(* IEC 61131-3 sources: daoli-st-library/DL_Process (part 5) *)

(* ---- FB_DL_PackMlUnitMode.st ---- *)
(*
  ==================================================================
  组件名 Component  : FB_DL_PackMlUnitMode
  分类   Category   : DL_Process
  版本   Version    : 1.0.1
  功能   Purpose    : PackML UnitMode 与 PMODE（PackML 状态模型）管理与命令过滤。
                      维护单元模式（生产 / 维护 / 手动 / 换型 / 清洗）与 PackML 状态
                      子集（空闲 / 启动 / 执行 / 保持 / 暂停 / 停止 / 中止 / 清除 /
                      复位 / 完成），按「当前状态 × 当前模式」两张闸对命令做过滤：
                      合法命令被受理并驱动状态迁移，非法命令被拒绝并给出拒绝原因；
                      模式切换仅在空闲 / 停止 / 完成三态允许。
  溯源   Origin     : PackML 状态与 UnitMode 组织为 OMAC PackML 公开标准语义；本件为
                      clean-room 实现，仅借鉴来源分类与参数域组织（来源标签
                      t2-7-packml 的 PackML 状态组织），未复制任何闭源代码行。
  平台   Platform   : 纯 IEC 61131-3（TON / R_TRIG / 枚举比较，无私有库）
  作者   Author     : 道莅代码库 · PLC 编程专家（R55）
  ------------------------------------------------------------------
  边界 Boundary     :
                      一 本件只做模式与状态管理及命令过滤，不执行任何设备动作（属主边界）；
                      二 中止（Abort）与停止（Stop）在全部模式下恒受理（安全侧优先）；
                      三 过渡态（启动 / 保持 / 暂停 / 停止 / 中止 / 清除 / 复位）由外部
                         完成信号 bTransDone 推进，并有过渡超时保护；
                      四 模式切换只在 eIdle / eStopped / eComplete 三态允许，其余态拒绝并留因；
                      五 无全局变量、无外部变量声明、无物理地址寻址。
  输出契约 Output contract:
                      eState / eMode 为锁存状态，只在合法迁移或合法模式切换时改变；
                      bCmdAccepted 为单拍脉冲（内部位置位、统一出口映射后撤销）；
                      eReject 每次拒绝独立留痕，nRejectCnt 饱和累计；
                      eCause 故障级成因与 bError 配对（R45），信息级永不置 bError。
  修订记录 Revision  :
    2026-11-20  v1.0.0  R55 首版（批 4 · 序号 19）
    2026-11-20  v1.0.1  R56 返修（7.5）：段 4 模式受理前补 eModeReq 枚举五选一合法性
                        校验，非法请求改记 eModeBlocked 不采纳（消除一拍非法模式窗口）；
                        段 9 / 段 10 头注释段号回正（原误标 segment 10 / 11）。
  ==================================================================
*)

TYPE E_DL_PmlState :
(
    eIdle        := 0,   // 空闲：允许启动与模式切换 / idle, start and mode change allowed
    eStarting    := 10,  // 启动过渡 / starting transition
    eExecute     := 20,  // 执行 / execute
    eCompleting  := 30,  // 完成过渡 / completing transition
    eComplete    := 40,  // 已完成：允许复位与模式切换 / complete, reset and mode change allowed
    eHolding     := 50,  // 保持过渡 / holding transition
    eHeld        := 60,  // 已保持 / held
    eUnholding   := 70,  // 解除保持过渡 / unholding transition
    eSuspending  := 80,  // 暂停过渡 / suspending transition
    eSuspended   := 90,  // 已暂停 / suspended
    eUnsuspending:= 100, // 解除暂停过渡 / unsuspending transition
    eStopping    := 110, // 停止过渡 / stopping transition
    eStopped     := 120, // 已停止：允许复位与模式切换 / stopped, reset and mode change allowed
    eClearing    := 130, // 清除过渡 / clearing transition
    eAborting    := 140, // 中止过渡 / aborting transition
    eAborted     := 150  // 已中止：只能经清除与复位恢复 / aborted, only clear and reset recover it
);
END_TYPE

TYPE E_DL_UnitMode :
(
    eProduction  := 0,   // 生产模式：全命令集 / production mode with the full command set
    eMaintenance := 10,  // 维护模式：禁暂停 / maintenance mode without suspend
    eManual      := 20,  // 手动模式：禁启动与保持 / manual mode without start and hold
    eChangeover  := 30,  // 换型模式：禁暂停与完成 / changeover mode without suspend and complete
    eCleaning    := 40   // 清洗模式：仅启动 / cleaning mode with start only
);
END_TYPE

TYPE E_DL_PmlCmd :
(
    eNone     := 0,      // 无命令 / no command
    eStart    := 10,     // 启动 / start
    eHold     := 20,     // 保持 / hold
    eUnhold   := 30,     // 解除保持 / unhold
    eSuspend  := 40,     // 暂停 / suspend
    eUnsuspend:= 50,     // 解除暂停 / unsuspend
    eStop     := 60,     // 停止 / stop
    eAbort    := 70,     // 中止 / abort
    eClear    := 80,     // 清除 / clear
    eReset    := 90,     // 复位 / reset
    eComplete := 100     // 完成 / complete
);
END_TYPE

TYPE E_DL_PmlReject :
(
    eNone            := 0, // 无拒绝 / no rejection
    eNoCmd           := 10, // 本拍无命令 / no command in this scan
    eIllegalState    := 20, // 该状态不接受此命令 / the current state does not accept this command
    eModeBlocked     := 30, // 当前模式禁止此命令 / the current mode blocks this command
    eModeLocked      := 40, // 当前状态不允许切换模式 / the current state does not allow a mode change
    eTransTimeout    := 50  // 过渡超时（故障级，与 bError 配对）/ transition timeout, a fault paired with bError
);
END_TYPE

FUNCTION_BLOCK FB_DL_PackMlUnitMode
VAR_INPUT
    bEnable      : BOOL := TRUE;             // 使能，失能时不受理命令并回空闲 [-] / enable, no command is accepted when disabled and the state returns to idle
    bReset       : BOOL := FALSE;           // 复位上升沿清故障锁存并回空闲 [-] / reset rising edge clears the fault latch and returns to idle
    bCmdStrobe   : BOOL := FALSE;            // 命令选通脉冲，上升沿消费 eCmdReq [-] / command strobe, eCmdReq is consumed on the rising edge
    eCmdReq      : E_DL_PmlCmd := E_DL_PmlCmd.eNone;   // 命令请求 [枚举] / requested command [enum]
    bModeStrobe  : BOOL := FALSE;            // 模式切换选通脉冲，上升沿消费 eModeReq [-] / mode change strobe, eModeReq is consumed on the rising edge
    eModeReq     : E_DL_UnitMode := E_DL_UnitMode.eProduction; // 模式请求 [枚举] / requested unit mode [enum]
    bTransDone   : BOOL := FALSE;            // 过渡完成信号（外部动作已完成）[-] / transition done signal from the external action
    tTransTo     : TIME := T#60S;            // 过渡超时 [毫秒]，域 大于零 / transition timeout [millisecond], domain above zero
END_VAR
VAR_OUTPUT
    eState       : E_DL_PmlState := E_DL_PmlState.eIdle;     // PackML 状态出口 [枚举] / PackML state outlet [enum]
    eMode        : E_DL_UnitMode := E_DL_UnitMode.eProduction; // 单元模式出口 [枚举] / unit mode outlet [enum]
    eAccepted    : E_DL_PmlCmd := E_DL_PmlCmd.eNone;         // 最近受理命令 [枚举] / last accepted command [enum]
    eReject      : E_DL_PmlReject := E_DL_PmlReject.eNone;   // 本拍拒绝原因 [枚举] / rejection reason of this scan [enum]
    bCmdAccepted : BOOL := FALSE;            // 命令受理单拍脉冲 [-] / command accepted single-shot pulse
    bModeAllowed : BOOL := FALSE;            // 当前状态是否允许切换模式 [-] / whether the current state allows a mode change
    bTransBusy   : BOOL := FALSE;            // 处于过渡态 [-] / inside a transition state
    uRejectCnt   : UDINT := 0;               // 拒绝计数（饱和到上限）[次] / rejection count, saturated [count]
    eCause       : E_DL_PmlReject := E_DL_PmlReject.eNone;   // 成因出口（复用拒绝枚举，故障级与 bError 配对）/ cause outlet reusing the reject enum, fault grade paired with bError
    bError       : BOOL := FALSE;            // 故障锁存标志 [-] / fault latch flag
END_VAR
VAR
    rtStrobe     : R_TRIG;                   // 命令选通沿检测，段 0 无条件刷新 / command strobe edge detector, refreshed unconditionally in segment zero
    rtMode       : R_TRIG;                   // 模式选通沿检测，段 0 无条件刷新 / mode strobe edge detector, refreshed unconditionally in segment zero
    rtReset      : R_TRIG;                   // 复位沿检测，段 0 无条件刷新 / reset edge detector, refreshed unconditionally in segment zero
    tonTrans     : TON;                      // 过渡超时，段 0 无条件刷新 / transition timeout, refreshed unconditionally in segment zero
    _eState      : E_DL_PmlState := E_DL_PmlState.eIdle;     // 内部状态，CASE 唯一写入目标 / internal state, the only CASE write target
    _eMode       : E_DL_UnitMode := E_DL_UnitMode.eProduction; // 内部模式锁存 / internal mode latch
    _eReject     : E_DL_PmlReject := E_DL_PmlReject.eNone;   // 本拍拒绝原因工作值 / rejection reason working value
    _eAccepted   : E_DL_PmlCmd := E_DL_PmlCmd.eNone;         // 本拍受理命令工作值（出口映射源）[枚举] / accepted command working value, source of the outlet [enum]
    _bFault      : BOOL := FALSE;            // 故障锁存位 [-] / fault latch bit
    _bInit       : BOOL := FALSE;            // 首扫初始化完成标志（R310）/ first scan initialisation flag
    _bAccInt     : BOOL := FALSE;            // 受理脉冲内部位，统一出口映射 / internal accepted bit, mapped at the unified outlet
    _bAccepted   : BOOL := FALSE;            // 本拍是否受理了命令 [-] / whether a command was accepted this scan
    _bTransBusy  : BOOL := FALSE;            // 过渡态判定 [-] / transition state verdict
    _bModeAllowed: BOOL := FALSE;            // 模式切换许可 [-] / mode change permission
    _bAllowStart : BOOL := FALSE;            // 模式允许启动 [-] / the mode allows start
    _bAllowHold  : BOOL := FALSE;            // 模式允许保持 [-] / the mode allows hold
    _bAllowSusp  : BOOL := FALSE;            // 模式允许暂停 [-] / the mode allows suspend
    _bAllowCompl : BOOL := FALSE;            // 模式允许完成 [-] / the mode allows complete
    _bModeValid  : BOOL := FALSE;            // 模式枚举合法 [-] / the mode enumeration is legal
    _bModeReqOk  : BOOL := FALSE;            // 模式请求枚举五选一合法性 [-] / whether the requested mode is one of the five legal members
    _uReject     : UDINT := 0;               // 拒绝计数工作值 [次] / rejection count working value [count]
END_VAR
VAR CONSTANT
    DL_PML_REJ_MAX : UDINT := 2000000000;    // 拒绝计数饱和上限（常量在 DINT 可表范围内）[次] / rejection count saturation ceiling, the constant fits in DINT
END_VAR

// 段 0｜定时器与沿检测无条件周期刷新（禁入分支），IN 只串过渡态闸 / segment 0, unconditional refresh with the transition gate on IN only
rtStrobe(CLK := bCmdStrobe); // 命令选通沿无条件刷新 / unconditional refresh of the command strobe
rtMode(CLK := bModeStrobe); // 模式选通沿无条件刷新 / unconditional refresh of the mode strobe
rtReset(CLK := bReset); // 复位沿无条件刷新 / unconditional refresh of the reset edge
tonTrans(IN := _bTransBusy AND (NOT _bFault) AND bEnable, PT := tTransTo); // 过渡超时，仅在过渡态计时 / transition timeout timing only inside a transition state

// 段 1｜首扫初始化（R310）/ segment 1, first scan initialisation
IF NOT _bInit THEN // 首扫一拍 / the very first scan
    _bInit := TRUE; // 置首扫完成标志 / raise the first scan flag
    _eState := E_DL_PmlState.eIdle; // 状态从空闲起步 / the state starts at idle
    _eMode := E_DL_UnitMode.eProduction; // 模式从生产起步 / the mode starts at production
    _eReject := E_DL_PmlReject.eNone; // 拒绝原因清零 / clear the rejection reason
    _bFault := FALSE; // 故障锁存清零 / clear the fault latch
    _uReject := 0; // 拒绝计数清零 / clear the rejection count
END_IF

// 段 2｜复位沿作用域：清锁存 / 迁状态 / 清脉冲内部位（模式保持，避免复位改工艺模式）/ segment 2, reset edge scope
IF rtReset.Q THEN // 复位沿 / reset edge
    _bFault := FALSE; // 作用域一：清故障锁存 / scope one, clear the fault latch
    _eReject := E_DL_PmlReject.eNone; // 作用域一：清拒绝原因 / scope one, clear the rejection reason
    _eState := E_DL_PmlState.eIdle; // 作用域二：迁回空闲 / scope two, migrate back to idle
    _bAccInt := FALSE; // 作用域二：清受理脉冲内部位 / scope two, clear the internal accepted bit
END_IF

// 段 3｜模式合法性与模式命令白名单（模式闸） / segment 3, mode validity and the per mode command whitelist
_bModeValid := (_eMode = E_DL_UnitMode.eProduction) OR (_eMode = E_DL_UnitMode.eMaintenance) OR (_eMode = E_DL_UnitMode.eManual) OR (_eMode = E_DL_UnitMode.eChangeover) OR (_eMode = E_DL_UnitMode.eCleaning); // 模式枚举五选一 / the mode is one of five
IF NOT _bModeValid THEN // 模式非法 / the mode is illegal
    _eMode := E_DL_UnitMode.eProduction; // 两级回退（R117）：一级回生产模式 / stage one of the two stage fallback, back to production
END_IF
_bAllowStart := (_eMode = E_DL_UnitMode.eProduction) OR (_eMode = E_DL_UnitMode.eMaintenance) OR (_eMode = E_DL_UnitMode.eChangeover) OR (_eMode = E_DL_UnitMode.eCleaning); // 启动白名单：手动模式禁启动 / start whitelist, manual mode forbids start
_bAllowHold := (_eMode = E_DL_UnitMode.eProduction) OR (_eMode = E_DL_UnitMode.eMaintenance) OR (_eMode = E_DL_UnitMode.eChangeover); // 保持白名单：手动与清洗禁保持 / hold whitelist, manual and cleaning forbid hold
_bAllowSusp := (_eMode = E_DL_UnitMode.eProduction); // 暂停白名单：仅生产模式 / suspend whitelist, production only
_bAllowCompl := (_eMode = E_DL_UnitMode.eProduction); // 完成白名单：仅生产模式 / complete whitelist, production only
_bModeAllowed := (_eState = E_DL_PmlState.eIdle) OR (_eState = E_DL_PmlState.eStopped) OR (_eState = E_DL_PmlState.eComplete); // 模式切换许可：空闲 / 停止 / 完成三态 / mode change allowed in idle, stopped and complete only

// 段 4｜模式切换：许可态内受理，非许可态留拒绝原因 / segment 4, mode change acceptance with a rejection trail
_eReject := E_DL_PmlReject.eNone; // 本拍拒绝原因预置空 / preset the rejection reason to none
_bModeReqOk := (eModeReq = E_DL_UnitMode.eProduction) OR (eModeReq = E_DL_UnitMode.eMaintenance) OR (eModeReq = E_DL_UnitMode.eManual) OR (eModeReq = E_DL_UnitMode.eChangeover) OR (eModeReq = E_DL_UnitMode.eCleaning); // 模式请求枚举五选一判式（R56 返修补齐）/ the requested mode is one of five legal members
IF rtMode.Q THEN // 模式选通沿 / mode strobe edge
    IF NOT bEnable THEN // 失能 / disabled
        _eReject := E_DL_PmlReject.eModeLocked; // 拒绝原因：失能不受理 / rejection reason, disabled
    ELSIF NOT _bModeReqOk THEN // 模式请求枚举非法 / the requested mode is illegal
        _eReject := E_DL_PmlReject.eModeBlocked; // 拒绝原因：非法模式请求不采纳（R56 返修补齐，消除一拍非法模式窗口）/ rejection reason, an illegal mode request is not adopted
    ELSIF _bModeAllowed THEN // 许可态 / inside a permitted state
        _eMode := eModeReq; // 采纳请求模式 / adopt the requested mode
    ELSE // 非许可态 / outside a permitted state
        _eReject := E_DL_PmlReject.eModeLocked; // 拒绝原因：状态锁模式 / rejection reason, the state locks the mode
    END_IF
END_IF

// 段 5｜过渡态判定 / segment 5, transition state verdict
_bTransBusy := (_eState = E_DL_PmlState.eStarting) OR (_eState = E_DL_PmlState.eCompleting) OR (_eState = E_DL_PmlState.eHolding) OR (_eState = E_DL_PmlState.eUnholding) OR (_eState = E_DL_PmlState.eSuspending) OR (_eState = E_DL_PmlState.eUnsuspending) OR (_eState = E_DL_PmlState.eStopping) OR (_eState = E_DL_PmlState.eClearing) OR (_eState = E_DL_PmlState.eAborting); // 九个过渡态之一 / one of the nine transition states

// 段 6｜过渡推进：外部完成信号或过渡超时（超时即中止并留故障级原因）/ segment 6, transition advancement by the external signal or by a timeout
IF _bTransBusy THEN // 过渡态内 / inside a transition state
    IF bTransDone THEN // 外部动作完成 / the external action completed
        CASE _eState OF
        E_DL_PmlState.eStarting: // 启动过渡完成 / starting completed
            _eState := E_DL_PmlState.eExecute; // 进执行态 / enter execute
        E_DL_PmlState.eCompleting: // 完成过渡完成 / completing completed
            _eState := E_DL_PmlState.eComplete; // 进已完成态 / enter complete
        E_DL_PmlState.eHolding: // 保持过渡完成 / holding completed
            _eState := E_DL_PmlState.eHeld; // 进已保持态 / enter held
        E_DL_PmlState.eUnholding: // 解除保持过渡完成 / unholding completed
            _eState := E_DL_PmlState.eExecute; // 回执行态 / back to execute
        E_DL_PmlState.eSuspending: // 暂停过渡完成 / suspending completed
            _eState := E_DL_PmlState.eSuspended; // 进已暂停态 / enter suspended
        E_DL_PmlState.eUnsuspending: // 解除暂停过渡完成 / unsuspending completed
            _eState := E_DL_PmlState.eExecute; // 回执行态 / back to execute
        E_DL_PmlState.eStopping: // 停止过渡完成 / stopping completed
            _eState := E_DL_PmlState.eStopped; // 进已停止态 / enter stopped
        E_DL_PmlState.eClearing: // 清除过渡完成 / clearing completed
            _eState := E_DL_PmlState.eIdle; // 回空闲态 / back to idle
        E_DL_PmlState.eAborting: // 中止过渡完成 / aborting completed
            _eState := E_DL_PmlState.eAborted; // 进已中止态 / enter aborted
        ELSE // 非法过渡态兜底（R128）/ illegal transition fallback
            _eState := E_DL_PmlState.eIdle; // 回空闲态 / back to idle
        END_CASE
    ELSIF tonTrans.Q THEN // 过渡超时 / the transition timed out
        _eReject := E_DL_PmlReject.eTransTimeout; // 故障级原因（与 bError 配对，R45）/ fault grade reason paired with bError
        _bFault := TRUE; // 置故障锁存 / raise the fault latch
        _eState := E_DL_PmlState.eAborting; // 强制走中止过渡 / force the aborting transition
    END_IF
END_IF

// 段 7｜命令过滤：状态闸在前、模式闸在后，两闸顺序固定（先判状态可接受性，再判模式白名单）/ segment 7, command filtering with the state gate before the mode gate
_eAccepted := E_DL_PmlCmd.eNone; // 受理命令预置空 / preset the accepted command to none
_bAccepted := FALSE; // 受理标志预置假 / preset the accepted flag to false
IF rtStrobe.Q AND bEnable AND (NOT _bFault) AND (NOT _bTransBusy) THEN // 选通沿、使能、无故障、非过渡态 / strobe while enabled, unfaulted and outside a transition
    IF eCmdReq = E_DL_PmlCmd.eNone THEN // 无命令 / no command
        _eReject := E_DL_PmlReject.eNoCmd; // 拒绝原因：无命令 / rejection reason, no command
    ELSE
        // 段 7.1｜状态闸：按当前状态给出可接受的命令集合 / segment 7.1, the state gate defines the acceptable command set
        CASE _eState OF
        E_DL_PmlState.eIdle: // 空闲态：启动 / 中止 / 复位 / 清除 / 模式许可 / idle state
            IF eCmdReq = E_DL_PmlCmd.eStart THEN // 启动 / start
                IF _bAllowStart THEN // 模式允许 / the mode allows it
                    _eState := E_DL_PmlState.eStarting; // 迁启动过渡 / enter starting
                    _eAccepted := E_DL_PmlCmd.eStart; // 受理启动 / accept start
                    _bAccepted := TRUE; // 置受理标志 / raise the accepted flag
                ELSE
                    _eReject := E_DL_PmlReject.eModeBlocked; // 模式闸拒绝 / blocked by the mode gate
                END_IF
            ELSIF eCmdReq = E_DL_PmlCmd.eAbort THEN // 中止 / abort
                _eState := E_DL_PmlState.eAborting; // 迁中止过渡 / enter aborting
                _eAccepted := E_DL_PmlCmd.eAbort; // 受理中止 / accept abort
                _bAccepted := TRUE; // 置受理标志 / raise the accepted flag
            ELSIF eCmdReq = E_DL_PmlCmd.eReset THEN // 复位 / reset
                _eState := E_DL_PmlState.eClearing; // 空闲态的复位等价于清除 / a reset from idle behaves as clearing
                _eAccepted := E_DL_PmlCmd.eReset; // 受理复位 / accept reset
                _bAccepted := TRUE; // 置受理标志 / raise the accepted flag
            ELSIF eCmdReq = E_DL_PmlCmd.eClear THEN // 清除 / clear
                _eState := E_DL_PmlState.eClearing; // 迁清除过渡 / enter clearing
                _eAccepted := E_DL_PmlCmd.eClear; // 受理清除 / accept clearing
                _bAccepted := TRUE; // 置受理标志 / raise the accepted flag
            ELSE // 其它命令 / any other command
                _eReject := E_DL_PmlReject.eIllegalState; // 状态闸拒绝 / blocked by the state gate
            END_IF
        E_DL_PmlState.eExecute: // 执行态：保持 / 暂停 / 停止 / 完成 / 中止 / execute state
            IF eCmdReq = E_DL_PmlCmd.eHold THEN // 保持 / hold
                IF _bAllowHold THEN // 模式允许 / the mode allows it
                    _eState := E_DL_PmlState.eHolding; // 迁保持过渡 / enter holding
                    _eAccepted := E_DL_PmlCmd.eHold; // 受理保持 / accept hold
                    _bAccepted := TRUE; // 置受理标志 / raise the accepted flag
                ELSE
                    _eReject := E_DL_PmlReject.eModeBlocked; // 模式闸拒绝 / blocked by the mode gate
                END_IF
            ELSIF eCmdReq = E_DL_PmlCmd.eSuspend THEN // 暂停 / suspend
                IF _bAllowSusp THEN // 模式允许 / the mode allows it
                    _eState := E_DL_PmlState.eSuspending; // 迁暂停过渡 / enter suspending
                    _eAccepted := E_DL_PmlCmd.eSuspend; // 受理暂停 / accept suspend
                    _bAccepted := TRUE; // 置受理标志 / raise the accepted flag
                ELSE
                    _eReject := E_DL_PmlReject.eModeBlocked; // 模式闸拒绝 / blocked by the mode gate
                END_IF
            ELSIF eCmdReq = E_DL_PmlCmd.eComplete THEN // 完成 / complete
                IF _bAllowCompl THEN // 模式允许 / the mode allows it
                    _eState := E_DL_PmlState.eCompleting; // 迁完成过渡 / enter completing
                    _eAccepted := E_DL_PmlCmd.eComplete; // 受理完成 / accept complete
                    _bAccepted := TRUE; // 置受理标志 / raise the accepted flag
                ELSE
                    _eReject := E_DL_PmlReject.eModeBlocked; // 模式闸拒绝 / blocked by the mode gate
                END_IF
            ELSIF eCmdReq = E_DL_PmlCmd.eStop THEN // 停止（安全侧恒受理）/ stop, always accepted on the safety side
                _eState := E_DL_PmlState.eStopping; // 迁停止过渡 / enter stopping
                _eAccepted := E_DL_PmlCmd.eStop; // 受理停止 / accept stop
                _bAccepted := TRUE; // 置受理标志 / raise the accepted flag
            ELSIF eCmdReq = E_DL_PmlCmd.eAbort THEN // 中止（安全侧恒受理）/ abort, always accepted
                _eState := E_DL_PmlState.eAborting; // 迁中止过渡 / enter aborting
                _eAccepted := E_DL_PmlCmd.eAbort; // 受理中止 / accept abort
                _bAccepted := TRUE; // 置受理标志 / raise the accepted flag
            ELSE // 其它命令 / any other command
                _eReject := E_DL_PmlReject.eIllegalState; // 状态闸拒绝 / blocked by the state gate
            END_IF
        E_DL_PmlState.eHeld: // 已保持态：解除保持 / 停止 / 中止 / held state
            IF eCmdReq = E_DL_PmlCmd.eUnhold THEN // 解除保持 / unhold
                _eState := E_DL_PmlState.eUnholding; // 迁解除保持过渡 / enter unholding
                _eAccepted := E_DL_PmlCmd.eUnhold; // 受理解除保持 / accept unhold
                _bAccepted := TRUE; // 置受理标志 / raise the accepted flag
            ELSIF eCmdReq = E_DL_PmlCmd.eStop THEN // 停止 / stop
                _eState := E_DL_PmlState.eStopping; // 迁停止过渡 / enter stopping
                _eAccepted := E_DL_PmlCmd.eStop; // 受理停止 / accept stop
                _bAccepted := TRUE; // 置受理标志 / raise the accepted flag
            ELSIF eCmdReq = E_DL_PmlCmd.eAbort THEN // 中止 / abort
                _eState := E_DL_PmlState.eAborting; // 迁中止过渡 / enter aborting
                _eAccepted := E_DL_PmlCmd.eAbort; // 受理中止 / accept abort
                _bAccepted := TRUE; // 置受理标志 / raise the accepted flag
            ELSE // 其它命令 / any other command
                _eReject := E_DL_PmlReject.eIllegalState; // 状态闸拒绝 / blocked by the state gate
            END_IF
        E_DL_PmlState.eSuspended: // 已暂停态：解除暂停 / 停止 / 中止 / suspended state
            IF eCmdReq = E_DL_PmlCmd.eUnsuspend THEN // 解除暂停 / unsuspend
                _eState := E_DL_PmlState.eUnsuspending; // 迁解除暂停过渡 / enter unsuspending
                _eAccepted := E_DL_PmlCmd.eUnsuspend; // 受理解除暂停 / accept unsuspend
                _bAccepted := TRUE; // 置受理标志 / raise the accepted flag
            ELSIF eCmdReq = E_DL_PmlCmd.eStop THEN // 停止 / stop
                _eState := E_DL_PmlState.eStopping; // 迁停止过渡 / enter stopping
                _eAccepted := E_DL_PmlCmd.eStop; // 受理停止 / accept stop
                _bAccepted := TRUE; // 置受理标志 / raise the accepted flag
            ELSIF eCmdReq = E_DL_PmlCmd.eAbort THEN // 中止 / abort
                _eState := E_DL_PmlState.eAborting; // 迁中止过渡 / enter aborting
                _eAccepted := E_DL_PmlCmd.eAbort; // 受理中止 / accept abort
                _bAccepted := TRUE; // 置受理标志 / raise the accepted flag
            ELSE // 其它命令 / any other command
                _eReject := E_DL_PmlReject.eIllegalState; // 状态闸拒绝 / blocked by the state gate
            END_IF
        E_DL_PmlState.eComplete: // 已完成态：复位 / 停止 / 中止 / complete state
            IF (eCmdReq = E_DL_PmlCmd.eReset) OR (eCmdReq = E_DL_PmlCmd.eClear) THEN // 复位或清除 / reset or clear
                _eState := E_DL_PmlState.eClearing; // 迁清除过渡 / enter clearing
                _eAccepted := eCmdReq; // 受理该命令 / accept that command
                _bAccepted := TRUE; // 置受理标志 / raise the accepted flag
            ELSIF eCmdReq = E_DL_PmlCmd.eAbort THEN // 中止 / abort
                _eState := E_DL_PmlState.eAborting; // 迁中止过渡 / enter aborting
                _eAccepted := E_DL_PmlCmd.eAbort; // 受理中止 / accept abort
                _bAccepted := TRUE; // 置受理标志 / raise the accepted flag
            ELSE // 其它命令 / any other command
                _eReject := E_DL_PmlReject.eIllegalState; // 状态闸拒绝 / blocked by the state gate
            END_IF
        E_DL_PmlState.eStopped: // 已停止态：复位 / 清除 / 中止 / stopped state
            IF (eCmdReq = E_DL_PmlCmd.eReset) OR (eCmdReq = E_DL_PmlCmd.eClear) THEN // 复位或清除 / reset or clear
                _eState := E_DL_PmlState.eClearing; // 迁清除过渡 / enter clearing
                _eAccepted := eCmdReq; // 受理该命令 / accept that command
                _bAccepted := TRUE; // 置受理标志 / raise the accepted flag
            ELSIF eCmdReq = E_DL_PmlCmd.eAbort THEN // 中止 / abort
                _eState := E_DL_PmlState.eAborting; // 迁中止过渡 / enter aborting
                _eAccepted := E_DL_PmlCmd.eAbort; // 受理中止 / accept abort
                _bAccepted := TRUE; // 置受理标志 / raise the accepted flag
            ELSE // 其它命令 / any other command
                _eReject := E_DL_PmlReject.eIllegalState; // 状态闸拒绝 / blocked by the state gate
            END_IF
        E_DL_PmlState.eAborted: // 已中止态：只能清除后复位 / aborted state, clear then reset only
            IF eCmdReq = E_DL_PmlCmd.eClear THEN // 清除 / clear
                _eState := E_DL_PmlState.eClearing; // 迁清除过渡 / enter clearing
                _eAccepted := E_DL_PmlCmd.eClear; // 受理清除 / accept clearing
                _bAccepted := TRUE; // 置受理标志 / raise the accepted flag
            ELSE // 其它命令 / any other command
                _eReject := E_DL_PmlReject.eIllegalState; // 状态闸拒绝 / blocked by the state gate
            END_IF
        ELSE // 过渡态不接受新命令 / transition states reject new commands
            _eReject := E_DL_PmlReject.eIllegalState; // 状态闸拒绝 / blocked by the state gate
        END_CASE
    END_IF
ELSIF rtStrobe.Q THEN // 有选通但使能 / 故障 / 过渡态不满足 / a strobe arrived under a blocking condition
    _eReject := E_DL_PmlReject.eIllegalState; // 拒绝原因：条件不满足 / rejection reason, the condition is not met
END_IF

// 段 8｜拒绝计数与受理脉冲内部位 / segment 8, rejection counting and the internal accepted bit
IF NOT (_eReject = E_DL_PmlReject.eNone) THEN // 本拍存在拒绝 / a rejection occurred
    IF _uReject < DL_PML_REJ_MAX THEN // 未达饱和上限 / below the ceiling
        _uReject := _uReject + 1; // 拒绝计数递增 / increment the rejection count
    END_IF
END_IF
IF _bAccepted THEN // 本拍受理了命令 / a command was accepted
    _bAccInt := TRUE; // 受理脉冲内部位置位（统一出口映射，R187）/ raise the internal accepted bit, mapped at the unified outlet
END_IF

// 段 9｜失能语义：不受理命令，状态保持但过渡计时停摆（R191 显式声明）/ segment 9, disabled semantics
IF NOT bEnable THEN // 失能 / disabled
    _bAccInt := FALSE; // 撤受理脉冲内部位 / withdraw the internal accepted bit
    _eReject := E_DL_PmlReject.eModeLocked; // 拒绝原因记模式锁（失能态不支持任何命令）/ rejection reason, disabled blocks every command
END_IF

// 段 10｜统一出口 / segment 10, unified outlet
eState := _eState; // 状态出口单点映射 / single-point state outlet mapping
eMode := _eMode; // 模式出口（锁存量）/ mode outlet from the latch
eAccepted := _eAccepted; // 受理命令出口 / accepted command outlet
eReject := _eReject; // 拒绝原因出口 / rejection reason outlet
bCmdAccepted := _bAccInt; // 受理脉冲映射本拍值 / map the accepted pulse for this scan
_bAccInt := FALSE; // 映射后立即撤销，保证单拍宽度（R187 两段式）/ revoke right after mapping to keep a single-scan width
bModeAllowed := _bModeAllowed; // 模式切换许可出口 / mode change permission outlet
bTransBusy := _bTransBusy; // 过渡态出口 / transition state outlet
uRejectCnt := _uReject; // 拒绝计数出口 / rejection count outlet
eCause := _eReject; // 成因出口与拒绝原因同源（名实双出口，R191）/ the cause outlet shares the rejection source
bError := _bFault; // 故障标志与锁存位同源 / the fault flag shares the latch source
END_FUNCTION_BLOCK

(* ---- FB_DL_PollTempBank.st ---- *)
(*==============================================================================
 * 组件名称 (Component)  : FB_DL_PollTempBank
 * 所属子库 (Sublibrary) : DL_Process
 * 当前版本 (Version)    : 1.0.0
 * 组件分类 (Category)   : 功能块（FUNCTION_BLOCK）· 工艺采集 · 温控器轮询采集行
 * 兼容性   (Platform)   : CODESYS 3.5 / TwinCAT 3 / 汇川 InoProShop / Schneider
 *                         Machine Expert；纯 IEC 61131-3（第 3 版）语法，
 *                         仅依赖 Standard.library（R_TRIG）
 * 功能描述 (Function)   : 一条温控器采集行——对最多 8 台温控器轮询采集过程值与设定值，
 *                         做工程量换算、有效域判定、滑动均值、偏差与最差通道定位，
 *                         输出通道质量掩码与在线台数，连续失败通道自动摘除并自动恢复。
 * 分层声明 (Layering)   : ① 调度归既有轮询主站件（本件内嵌其一个实例，只注入站表与
 *                         节拍参数，不重写调度、重试与超时逻辑）；② 滤波归既有滑动均值件
 *                         （本件为八个通道各持一个实例，只给样本与采样允许）；
 *                         ③ 本件只做「行级编排加通道质量」，不做温控闭环——设定值下发、
 *                         自整定、超温切断属温控器内部或工艺层职责，本件只读不写。
 * 传输层说明 (Transport) : 内嵌的调度实例以库内基类形态声明，其帧收发为抽象桩。生产部署
 *                         时必须由具备真实串口或网口收发的派生块替换该声明，否则调度层会
 *                         锁「传输层未实现」故障、全部通道因轮询不成功而逐台摘除。这一
 *                         失败是**可观测的显式失败**（质量掩码全置位、在线台数为零），
 *                         不会静默给出假温度，故不在本件内把它翻译成故障码。
 * 保持策略 (Hold)       : 坏通道的温度保持上次有效值并在质量掩码里标记，**绝不**用零或
 *                         上限值填充——零摄氏度在锂电烘箱、冷库等场景是合法工况值，用零
 *                         填充会掩盖真实故障（与既有温度扫描件同一纪律）。
 * 摘除与恢复 (Drop)     : 连续失败达到阈值即摘除并置信息码；摘除后仍继续轮询该通道，
 *                         连续两拍有效即自动恢复。若不继续轮询，被摘除的通道永远拿不到
 *                         有效数据、也就永远无法恢复，这是摘除策略必须配对的另一半。
 * 职责边界 (Scope)      : 不做写设定值（只采集）、不做地址表编辑器的校验（站表按默认值
 *                         填充，机型差异由调用方改表）、不做历史归档与报警分级。
 * 开源溯源 (Origin)     : 来源标签 roadmap-p0 加 t1-4。原创实现（参考 ROADMAP §13.6 P0
 *                         条目「温控器轮询采集行（复用轮询主站与滑动均值）」的需求定义，
 *                         以及 CODESYS Forge ModbusFB 族「调度与传输分层」的组织方式）。
 *                         仅借组织方式与参数域，编排逻辑、通道质量掩码、摘除与恢复策略、
 *                         枚举、状态机与全部码位 100% 本库独立设计，clean-room 实现，
 *                         不复制任何示例代码与注释。
 * 依赖     (Depends)    : ST_DL_PollItem 与 FB_DL_ModbusPollMaster（DL_Process 既有件，
 *                         本件只引用不声明）；FB_DL_MovingAverage（DL_MathData 既有件）；
 *                         Standard.library: R_TRIG
 * 故障码表 (Error codes):
 *   16#0005_0108【信息级】台数、窗口长度或摘除阈值越界已钳位
 *   16#0005_0109【信息级】通道连续失败达到阈值已摘除（仍继续轮询以便自动恢复）
 *   16#0005_010A【信息级】滤波窗口为 1，均值等于瞬时值（无滤波能力）
 *   16#0005_0207【故障级】换算比例非正，量纲错且含零乘隐患（锁存）
 *   16#0005_0208【故障级】有效温度域为空，任何读数都会被判无效（锁存）
 *   16#0005_0209【故障级】非法状态兜底（锁存，终端安全态）
 * 码位占用 (Slot)       : 信息级 0108 / 0109 / 010A；故障级 0207 / 0208 / 0209。
 *                         全部落在 R12 本件分配块内，无跨块借用、无段外哨兵值。
 * 拍序纪律 (Cycle order) :
 *   ① ePhase        ：段 7 状态机（唯一位移点），段 8 复位分支是唯一回退点
 *   ② 三个生效参数   ：段 4 单点钳位，后续所有数组访问与循环上限都取这三个生效值
 *   ③ 质量掩码       ：段 6 装配后整值写出，与本拍在线台数、最差通道同拍一致
 *   ④ uErrorId       ：段 9 单一优先级链，全拍只写一次
 * 验收向量 (Acceptance) :
 *   V1 单台正常：台数 1、过程值 253、设定值 250、比例 0.1 → 温度 25.3、设定 25.0、
 *      偏差 0.3、质量掩码为零、在线 1 台
 *   V2 超域：第 2 台过程值 3200（换算 320.0 高于上限 200）→ 该通道无效、温度保持、
 *      质量掩码位 1 置位、连续失败计数 1
 *   V3 摘除：第 3 台连续三拍轮询失败、阈值为 3 → 第 3 拍摘除、质量掩码位 2 置位、
 *      在线台数减 1、码 0109
 *   V4 最差通道：两通道偏差分别负 3.5 与正 4.2 → 最差通道号为 4、最差偏差正 4.2
 *   V5 量纲错：比例为 0 → 故障位置位、码 0207、各通道温度保持
 * 偏离留档 (Deviation)  :
 *   ① 规格第 3.18 节正文提到「评估相」，但 §2.1 的枚举只有三成员。本件按枚举实现，
 *      把逐通道评估并入轮询相的固定段完成，不新增枚举成员，避免枚举与码表、文档三处
 *      不一致。
 *   ② 规格要求「内嵌调度实例」，但库内调度基类的传输层为抽象桩，无法在本文件内以派生块
 *      替换其声明。本件保留基类实例并在头注释写明部署要求，把「传输层未就绪」表现为
 *      质量掩码全坏这一可观测结果，而不是伪造成功。
 *   ③ 参数钳位放在状态机之前的固定段（而非待机相），理由：台数决定站表填充与循环上限，
 *      必须每拍先于任何数组访问生效，否则上电首拍会用未钳位值访问数组。
 * 修订历史 (Revision)   :
 *   2026-11-15  v1.0.0  首版落盘（R12 · 泳道 C · 温控器轮询采集行 P0 件）
 *============================================================================*)

(*------------------------------------------------------------------------------
 * 枚举: E_DL_TempBankPhase（本块相位，归属本功能块并同文件发布）
 *       Phase enumeration owned by this block
 *-----------------------------------------------------------------------------*)
TYPE E_DL_TempBankPhase :
(
    eIdle    := 0,   // 待机：未使能或参数闸门未过，输出保持 / Idle, disabled or the gate has not passed
    ePolling := 10,  // 轮询：调度实例推进轮询，同时做逐通道换算与质量判定 / Polling with per-channel evaluation
    eFault   := 99   // 故障：量纲错、有效域为空或非法状态，需复位退出 / Fault, needs a reset to leave
);
END_TYPE

FUNCTION_BLOCK FB_DL_PollTempBank
VAR_INPUT
    bEnable        : BOOL;                              // 使能，FALSE 时暂停轮询并保持输出 [-] / Enable, polling paused and outputs held while FALSE
    bReset         : BOOL;                              // 复位故障与摘除状态，上升沿有效 [-] / Rising edge clears the fault and the drop state
    nDeviceCount   : INT := 4;                          // 温控器台数 [台]，有效域 1 到 8 / Device count, one to eight
    anSlaveAddr    : ARRAY[1..8] OF USINT;              // 各台从站地址 [1 到 247] / Slave address per device
    auPvRaw        : ARRAY[1..8] OF INT;                // 各台过程值原始寄存器，由传输层写入 [原始码] / Raw process values written by the transport
    auSvRaw        : ARRAY[1..8] OF INT;                // 各台设定值原始寄存器 [原始码] / Raw setpoints
    abPollOk       : ARRAY[1..8] OF BOOL;               // 各台本次轮询成功标志 [-] / Per-device poll success flags
    fScaleGain     : REAL := 0.1;                       // 原始码到温度的比例 [摄氏度每码]，域大于 0 / Raw to temperature gain, must exceed zero
    fScaleOffset   : REAL := 0.0;                       // 零点偏移 [摄氏度] / Zero offset in degrees Celsius
    fRangeMin      : REAL := -50.0;                     // 有效温度下限 [摄氏度] / Valid temperature lower bound
    fRangeMax      : REAL := 200.0;                     // 有效温度上限 [摄氏度] / Valid temperature upper bound
    nFilterLen     : INT := 8;                          // 滑动均值窗口长度 [拍]，有效域 1 到 32 / Moving average window, one to thirty-two
    nDropAfterFails: INT := 3;                          // 连续失败多少次摘除通道 [次]，有效域 1 到 10 / Failures before dropping a channel
END_VAR
VAR_OUTPUT
    afTempC        : ARRAY[1..8] OF REAL;               // 各台温度 [摄氏度]，坏通道保持上次有效值 / Temperature per device, bad channels hold the last value
    afSetpointC    : ARRAY[1..8] OF REAL;               // 各台设定值 [摄氏度] / Setpoint per device
    afDeviation    : ARRAY[1..8] OF REAL;               // 各台偏差，过程值减设定值 [摄氏度] / Deviation, process minus setpoint
    afTempAvg      : ARRAY[1..8] OF REAL;               // 各台滑动均值 [摄氏度] / Per-device moving average
    auCommFailCnt  : ARRAY[1..8] OF UINT;               // 各台连续失败次数，饱和到上限 [次] / Consecutive failure counter per device, saturated
    uQualityMask   : WORD;                              // 通道坏质量掩码，位 n 减一 对应第 n 台 [位串] / Bad channel mask, bit n minus one is device n
    nOnlineCount   : INT;                               // 在线台数 [台] / Online device count
    nWorstIdx      : INT;                               // 偏差绝对值最大的在线通道号，0 表示无 [通道号] / Channel with the largest absolute deviation
    fWorstDev      : REAL;                              // 该通道的有符号偏差值 [摄氏度] / Signed deviation of that channel
    bError         : BOOL;                              // 故障级锁存，仅 0207 至 0209 置位 [-] / Latched fault, only fault level codes set it
    uErrorId       : UDINT;                             // 事件码，0 表示无事件 [代码] / Event code, zero means none
    eState         : E_DL_TempBankPhase;                // 主状态机当前相位 [-] / Current phase of the main state machine
END_VAR
VAR_IN_OUT
    aPollTable     : ARRAY[0..15] OF ST_DL_PollItem;    // 轮询站表，由内嵌调度实例持有并更新统计 [-] / Poll table owned by the embedded scheduler
END_VAR
VAR
    fbPoll         : FB_DL_ModbusPollMaster;            // 内嵌轮询调度实例，主周期无条件调用 / Embedded poll scheduler, called unconditionally
    afbAvg         : ARRAY[1..8] OF FB_DL_MovingAverage; // 逐通道滑动均值实例，主周期无条件全量调用 / Per-channel moving average instances
    fbTrigReset    : R_TRIG;                            // 复位沿检测，主周期无条件刷新 [-] / Reset edge detector, refreshed unconditionally
    ePhase         : E_DL_TempBankPhase := E_DL_TempBankPhase.eIdle; // 内部相位，对外经 eState 输出 [-] / Internal phase exported as eState
    bInit          : BOOL := FALSE;                     // 首扫标志，初值 FALSE，判据取非 [-] / First-scan flag initialised FALSE
    bFaultLatch    : BOOL;                              // 故障锁存，仅复位分支清除 [-] / Fault latch, cleared by the reset path only
    uErrInt        : UDINT;                             // 故障级码寄存，锁存型 [代码] / Latched fault level code register
    uInfoCode      : UDINT;                             // 本拍信息级码，每拍重算 [代码] / Info level code recomputed every scan
    nDevUse        : INT := 1;                          // 生效台数，钳位后 [台] / Effective device count after clamping
    nFilterUse     : INT := 1;                          // 生效窗口长度，钳位后 [拍] / Effective window length after clamping
    nDropUse       : INT := 1;                          // 生效摘除阈值，钳位后 [次] / Effective drop threshold after clamping
    fGainUse       : REAL := 1.0;                       // 生效换算比例 [摄氏度每码] / Effective gain
    bEval          : BOOL;                              // 本拍执行通道评估 [-] / Evaluation enabled flag of this scan
    bDropEvent     : BOOL;                              // 本拍有通道被摘除 [-] / A channel was dropped this scan
    fVal           : REAL;                              // 单通道温度 [摄氏度] / Single channel temperature
    fSp            : REAL;                              // 单通道设定值 [摄氏度] / Single channel setpoint
    fDevAbs        : REAL;                              // 偏差绝对值 [摄氏度] / Absolute deviation
    fWorstTmp      : REAL;                              // 最差偏差绝对值暂存 [摄氏度] / Worst absolute deviation temporary
    uQBuild        : WORD;                              // 质量掩码装配 [位串] / Quality mask under assembly
    nOnline        : INT;                               // 在线计数 [台] / Online counter
    nWorst         : INT;                               // 最差通道号 [通道号] / Worst channel number
    abOkTmp        : ARRAY[1..8] OF BOOL;               // 各通道本拍有效标志 [-] / Per-channel validity of this scan
    abDropped      : ARRAY[1..8] OF BOOL;               // 通道已摘除标志 [-] / Channel dropped flags
    anRecover      : ARRAY[1..8] OF INT;                // 摘除后连续有效拍数 [拍] / Consecutive valid scans after a drop
    bValFin        : BOOL;                              // 换算值有限标志 [-] / Finite converted value flag
    nGuard         : DINT;                              // 循环守卫计数 [次]，上限常量化 / Loop guard counter with a constant bound
    i              : INT;                               // 通道索引 [1..8] / Channel loop index
    k              : INT;                               // 站表索引 [0..15] / Poll table loop index
END_VAR
VAR CONSTANT
    DL_DEV_MAX     : INT := 8;                          // 温控器台数上限 [台] / Device count limit
    DL_FILT_MAX    : INT := 32;                         // 滤波窗口上限 [拍] / Window length limit
    DL_DROP_MAX    : INT := 10;                         // 摘除阈值上限 [次] / Drop threshold limit
    DL_TABLE_MAX   : INT := 16;                         // 站表长度 [项] / Poll table length
    DL_FAIL_MAX    : UINT := 9999;                      // 连续失败计数饱和值 [次] / Failure counter saturation
    DL_MASK_ONE    : WORD := 16#0001;                   // 单通道基准位 [位串] / Single channel base bit
    DL_MASK_NONE   : WORD := 16#0000;                   // 全零掩码基准 [位串] / All zero mask reference
    DL_GAIN_MIN    : REAL := 1.0E-6;                    // 比例最小正值 [摄氏度每码] / Minimum positive gain
    DL_GAIN_SAFE   : REAL := 1.0;                       // 比例非法时的兜底值 [摄氏度每码] / Safe gain used when the input is illegal
    DL_TEMP_MAX    : REAL := 1.0E6;                     // 温度量级上限，超出视为非有限 [摄氏度] / Temperature magnitude bound
    DL_GUARD_MAX   : DINT := 64;                        // 循环守卫上限 [次] / Loop guard bound
    DL_RECOVER_NEED: INT := 2;                          // 自动恢复所需的连续有效拍数 [拍] / Valid scans required for an automatic recovery
    DL_FUNC_READ   : USINT := 3;                        // 读保持寄存器功能码 [功能码] / Read holding registers function code
    DL_REG_QTY     : UINT := 2;                         // 每站连续读两个寄存器，过程值与设定值 [个] / Two registers per station
    DL_REG_START   : UINT := 0;                         // 站表起始地址 [寄存器地址] / Station start address
    DL_RESP_TO     : TIME := T#500MS;                   // 单事务响应超时 [毫秒] / Per-transaction response timeout
    DL_POLL_GAP    : TIME := T#50MS;                    // 相邻事务最小间隔 [毫秒] / Minimum poll interval
    DL_RETRY_MAX   : UINT := 2;                         // 超时重试上限 [次] / Retry limit
END_VAR

(*------------------------------------------------------------------------------
 * 段 1｜输出确定性默认值（单拍与评估缓冲每拍预清零，R25 第一律）
 *      Deterministic defaults first, evaluation buffers pre-cleared every scan
 *-----------------------------------------------------------------------------*)
uInfoCode  := 16#0000_0000;                     // 信息级码每拍重算（Info code recomputed every scan）
nGuard     := 0;                                // 循环守卫清零（Loop guard cleared）
bDropEvent := FALSE;                            // 摘除事件标志预清零（Drop event flag pre-cleared）
bEval      := bEnable AND (ePhase = E_DL_TempBankPhase.ePolling); // 评估使能取上一拍相位（Evaluation enabled from the previous phase）
FOR i := 1 TO DL_DEV_MAX DO
    abOkTmp[i] := FALSE;                        // 本拍有效标志预清零，未轮询时不采样（No sampling while the phase is not polling）
END_FOR

(*------------------------------------------------------------------------------
 * 段 2｜沿检测无条件刷新（红线：实例在 CASE 之外每拍必刷）
 *      Edge detection refreshed unconditionally outside the CASE
 *-----------------------------------------------------------------------------*)
fbTrigReset(CLK := bReset);

(*------------------------------------------------------------------------------
 * 段 3｜首扫初始化（唯一合法范式：初值 FALSE，判据取非）
 *      First-scan initialisation following the single legal pattern
 *-----------------------------------------------------------------------------*)
IF NOT bInit THEN
    FOR i := 1 TO DL_DEV_MAX DO
        afTempC[i]       := 0.0;                // 温度出口清零（Temperature outlet cleared）
        afSetpointC[i]   := 0.0;                // 设定值出口清零（Setpoint outlet cleared）
        afDeviation[i]   := 0.0;                // 偏差出口清零（Deviation outlet cleared）
        afTempAvg[i]     := 0.0;                // 均值出口清零（Average outlet cleared）
        auCommFailCnt[i] := 0;                  // 连续失败计数清零（Failure counter cleared）
        abDropped[i]     := FALSE;              // 摘除标志清零（Drop flag cleared）
        anRecover[i]     := 0;                  // 恢复计数清零（Recovery counter cleared）
    END_FOR
    uQualityMask := DL_MASK_NONE;               // 质量掩码清零（Quality mask cleared）
    nOnlineCount := 0;                          // 在线台数清零（Online count cleared）
    nWorstIdx    := 0;                          // 最差通道清零（Worst channel cleared）
    fWorstDev    := 0.0;                        // 最差偏差清零（Worst deviation cleared）
    nDevUse      := 1;                          // 生效台数取下限（Effective device count at the lower bound）
    nFilterUse   := 1;                          // 生效窗口取下限（Effective window at the lower bound）
    nDropUse     := 1;                          // 生效阈值取下限（Effective threshold at the lower bound）
    fGainUse     := DL_GAIN_SAFE;               // 生效比例取兜底值（Effective gain set to the safe value）
    bFaultLatch  := FALSE;                      // 故障锁存清零（Fault latch cleared）
    uErrInt      := 16#0000_0000;               // 故障码清零（Fault code cleared）
    ePhase       := E_DL_TempBankPhase.eIdle;   // 相位复位为待机（Phase reset to idle）
    bInit        := TRUE;                       // 首扫只做一次（First scan runs once）
END_IF

(*------------------------------------------------------------------------------
 * 段 4｜参数钳位（先于任何数组访问与循环上限；越界只钳位并置信息码）
 *      Parameter clamping before any array access or loop bound
 *-----------------------------------------------------------------------------*)
IF nDeviceCount < 1 THEN
    nDevUse   := 1;                             // 台数下限钳位（Clamped to the lower bound）
    uInfoCode := 16#0005_0108;                  // 0108 台数越界已钳位（Device count clamped）
ELSIF nDeviceCount > DL_DEV_MAX THEN
    nDevUse   := DL_DEV_MAX;                    // 台数上限钳位（Clamped to the upper bound）
    uInfoCode := 16#0005_0108;                  // 0108 台数越界已钳位（Device count clamped）
ELSE
    nDevUse   := nDeviceCount;                  // 合法台数直通（Valid device count passed through）
END_IF

IF nFilterLen < 1 THEN
    nFilterUse := 1;                            // 窗口下限钳位（Clamped to the lower bound）
    uInfoCode  := 16#0005_0108;                 // 0108 窗口越界已钳位（Window clamped）
ELSIF nFilterLen > DL_FILT_MAX THEN
    nFilterUse := DL_FILT_MAX;                  // 窗口上限钳位（Clamped to the upper bound）
    uInfoCode  := 16#0005_0108;                 // 0108 窗口越界已钳位（Window clamped）
ELSE
    nFilterUse := nFilterLen;                   // 合法窗口直通（Valid window passed through）
END_IF
IF nFilterUse = 1 THEN
    uInfoCode := 16#0005_010A;                  // 010A 窗口为 1，无滤波能力（Window of one gives no filtering）
END_IF

IF nDropAfterFails < 1 THEN
    nDropUse  := 1;                             // 阈值下限钳位（Clamped to the lower bound）
    uInfoCode := 16#0005_0108;                  // 0108 阈值越界已钳位（Threshold clamped）
ELSIF nDropAfterFails > DL_DROP_MAX THEN
    nDropUse  := DL_DROP_MAX;                   // 阈值上限钳位（Clamped to the upper bound）
    uInfoCode := 16#0005_0108;                  // 0108 阈值越界已钳位（Threshold clamped）
ELSE
    nDropUse  := nDropAfterFails;               // 合法阈值直通（Valid threshold passed through）
END_IF

IF fScaleGain <= DL_GAIN_MIN THEN
    fGainUse := DL_GAIN_SAFE;                   // 量纲错：兜底比例避免零乘（Safe gain avoids a zero product）
    IF NOT bFaultLatch THEN
        bFaultLatch := TRUE;                    // 锁故障，保留首出码（Latch the fault keeping the first code）
        uErrInt     := 16#0005_0207;            // 0207 换算比例非正（Non-positive gain）
    END_IF
ELSE
    fGainUse := fScaleGain;                     // 合法比例直通（Valid gain passed through）
END_IF

IF fRangeMin >= fRangeMax THEN
    IF NOT bFaultLatch THEN
        bFaultLatch := TRUE;                    // 有效域为空：锁故障（Empty valid range, latch the fault）
        uErrInt     := 16#0005_0208;            // 0208 有效域为空（Empty valid range）
    END_IF
END_IF

(*------------------------------------------------------------------------------
 * 段 5｜站表默认值填充与调度实例调用（实例每拍无条件调用，使能经引脚注入）
 *      Poll table defaults and the embedded scheduler, called every scan
 *-----------------------------------------------------------------------------*)
FOR k := 0 TO (DL_TABLE_MAX - 1) DO
    nGuard := nGuard + 1;                       // 守卫递增（Guard incremented）
    IF nGuard > DL_GUARD_MAX THEN
        EXIT;                                   // 守卫到顶即退出（Bail out at the guard bound）
    END_IF
    IF k < DL_DEV_MAX THEN
        IF (k + 1) <= nDevUse THEN
            aPollTable[k].uSlaveAddr := anSlaveAddr[k + 1]; // 从站地址取引脚（Slave address from the pin）
            aPollTable[k].uFuncCode  := DL_FUNC_READ;       // 读保持寄存器（Read holding registers）
            aPollTable[k].uStartAddr := DL_REG_START;       // 起始地址零（Start address zero）
            aPollTable[k].uQuantity  := DL_REG_QTY;         // 连续两寄存器：过程值与设定值（Two registers, process and setpoint）
            aPollTable[k].bSkip      := FALSE;              // 启用本站（Station enabled）
        ELSE
            aPollTable[k].bSkip := TRUE;                    // 超出台数：跳过（Beyond the device count, skip）
        END_IF
    ELSE
        aPollTable[k].bSkip := TRUE;                        // 站表多余项一律跳过（Extra table entries are skipped）
    END_IF
END_FOR

fbPoll(bEnable       := bEnable AND (ePhase = E_DL_TempBankPhase.ePolling),
       uStationCount := INT_TO_UINT(nDevUse),
       tRespTimeout  := DL_RESP_TO,
       uMaxRetry     := DL_RETRY_MAX,
       tPollInterval := DL_POLL_GAP,
       aPollTable    := aPollTable);            // 调度实例无条件调用，绝不做条件包裹（Never wrapped in a conditional）

(*------------------------------------------------------------------------------
 * 段 6｜逐通道评估（换算、三道有效性闸、失败计数与摘除、恢复、偏差与最差通道）
 *      Per-channel evaluation with the three validity gates and the drop policy
 *-----------------------------------------------------------------------------*)
IF bEval THEN
    nOnline     := 0;                           // 在线计数清零（Online counter cleared）
    nWorst      := 0;                           // 最差通道清零（Worst channel cleared）
    fWorstTmp   := 0.0;                         // 最差偏差暂存清零（Worst deviation temporary cleared）
    uQBuild     := DL_MASK_NONE;                // 质量掩码装配清零（Quality mask cleared）
    FOR i := 1 TO DL_DEV_MAX DO
        nGuard := nGuard + 1;                   // 守卫递增（Guard incremented）
        IF nGuard > DL_GUARD_MAX THEN
            EXIT;                               // 守卫到顶即退出（Bail out at the guard bound）
        END_IF
        IF i <= nDevUse THEN
            fVal    := (INT_TO_REAL(auPvRaw[i]) * fGainUse) + fScaleOffset; // 过程值换算（Process value conversion）
            fSp     := (INT_TO_REAL(auSvRaw[i]) * fGainUse) + fScaleOffset; // 设定值换算（Setpoint conversion）
            bValFin := NOT ((fVal <> fVal) OR (ABS(fVal) > DL_TEMP_MAX));   // 有限性判定（Finiteness test）
            abOkTmp[i] := abPollOk[i] AND bValFin AND (fVal >= fRangeMin) AND (fVal <= fRangeMax); // 三道闸（Three gates）
            IF abOkTmp[i] THEN
                auCommFailCnt[i] := 0;          // 有效拍清零连续失败（Clear the failure counter）
                afTempC[i]       := fVal;       // 有效才刷新温度（Refresh the temperature only when valid）
                afSetpointC[i]   := fSp;        // 有效才刷新设定值（Refresh the setpoint only when valid）
                IF abDropped[i] THEN
                    IF anRecover[i] < DL_RECOVER_NEED THEN
                        anRecover[i] := anRecover[i] + 1; // 恢复计数累加（Recovery counter incremented）
                    END_IF
                    IF anRecover[i] >= DL_RECOVER_NEED THEN
                        abDropped[i] := FALSE;  // 连续有效达阈值：自动恢复（Automatic recovery）
                        anRecover[i] := 0;      // 恢复计数清零（Recovery counter cleared）
                    END_IF
                END_IF
            ELSE
                IF auCommFailCnt[i] < DL_FAIL_MAX THEN
                    auCommFailCnt[i] := auCommFailCnt[i] + 1; // 连续失败累加，饱和到上限（Failure counter incremented and saturated）
                END_IF
                anRecover[i] := 0;              // 失败即清恢复计数（Recovery counter cleared on a failure）
                IF (NOT abDropped[i]) AND (auCommFailCnt[i] >= INT_TO_UINT(nDropUse)) THEN
                    abDropped[i] := TRUE;       // 达阈值：摘除通道（Drop the channel）
                    bDropEvent   := TRUE;       // 标记待置信息码 0109（Flag the informational code 0109）
                END_IF
            END_IF
            IF abDropped[i] OR (NOT abOkTmp[i]) THEN
                uQBuild := uQBuild OR SHL(DL_MASK_ONE, i - 1); // 坏通道进位（Bad channel bit set）
            ELSE
                nOnline := nOnline + 1;         // 在线台数累加（Online count incremented）
            END_IF
            afDeviation[i] := afTempC[i] - afSetpointC[i]; // 偏差由保持后的温度算出（Deviation from the held temperature）
            IF (NOT abDropped[i]) AND abOkTmp[i] THEN
                fDevAbs := ABS(afDeviation[i]);  // 只让在线通道参与最差判定（Only online channels compete）
                IF fDevAbs > fWorstTmp THEN
                    fWorstTmp := fDevAbs;        // 严格大于才替换，并列取小号（Strictly greater, ties keep the lower index）
                    nWorst    := i;              // 记录最差通道号（Record the worst channel）
                END_IF
            END_IF
        ELSE
            abOkTmp[i]     := FALSE;            // 超出台数：本拍无效（Beyond the device count, invalid）
            afDeviation[i] := 0.0;              // 超出台数：偏差清零（Deviation cleared）
        END_IF
    END_FOR
    uQualityMask := uQBuild;                    // 质量掩码整值写出（Quality mask published as a whole）
    nOnlineCount := nOnline;                    // 在线台数写出（Online count published）
    nWorstIdx    := nWorst;                     // 最差通道写出（Worst channel published）
    IF nWorst > 0 THEN
        fWorstDev := afDeviation[nWorst];       // 最差通道的有符号偏差（Signed deviation of that channel）
    ELSE
        fWorstDev := 0.0;                       // 无在线通道时为零（Zero when no channel is online）
    END_IF
    IF bDropEvent THEN
        uInfoCode := 16#0005_0109;              // 0109 通道已摘除（A channel was dropped）
    END_IF
END_IF

(*------------------------------------------------------------------------------
 * 段 7｜滑动均值实例全量调用（红线：实例每拍无条件调用，采样经允许位控制）
 *      Moving average instances called for every channel, sampling gated by a flag
 *-----------------------------------------------------------------------------*)
FOR i := 1 TO DL_DEV_MAX DO
    nGuard := nGuard + 1;                       // 守卫递增（Guard incremented）
    IF nGuard > DL_GUARD_MAX THEN
        EXIT;                                   // 守卫到顶即退出（Bail out at the guard bound）
    END_IF
    afbAvg[i](fInput      := afTempC[i],
              nWindowSize := nFilterUse,
              bSample     := bEval AND abOkTmp[i],
              bEnable     := TRUE,
              bReset      := fbTrigReset.Q);    // 复位沿同拍清窗口，避免复位后混旧样本（Reset clears the window）
    afTempAvg[i] := afbAvg[i].fAverage;         // 均值出口（Average outlet）
END_FOR

(*------------------------------------------------------------------------------
 * 段 8｜主状态机（枚举每个成员均有标签，末尾 ELSE 兜底到终端安全态）
 *      Main state machine, one label per member plus a trailing ELSE fallback
 *-----------------------------------------------------------------------------*)
CASE ePhase OF

    E_DL_TempBankPhase.eIdle: // 待机：故障或未使能则停留，否则进入轮询
        IF bFaultLatch THEN
            ePhase := E_DL_TempBankPhase.eFault;   // 参数已锁故障：进故障态（Gate failed, enter the fault state）
        ELSIF bEnable THEN
            ePhase := E_DL_TempBankPhase.ePolling; // 进轮询相（Enter the polling phase）
        END_IF

    E_DL_TempBankPhase.ePolling: // 轮询：评估在固定段完成，本相只负责相位迁移
        IF NOT bEnable THEN
            ePhase := E_DL_TempBankPhase.eIdle;    // 掉使能：回待机，输出保持（Disabled, back to idle with outputs held）
        ELSIF bFaultLatch THEN
            ePhase := E_DL_TempBankPhase.eFault;   // 运行期参数失效：进故障态（A parameter failed at run time）
        END_IF

    E_DL_TempBankPhase.eFault: // 故障：输出保持，等复位沿
        IF fbTrigReset.Q THEN
            ePhase := E_DL_TempBankPhase.eIdle;    // 复位后回待机，重新过闸门（Reset returns to idle and re-runs the gate）
        END_IF

    ELSE
        bFaultLatch := TRUE;                        // 非法状态兜底锁存（Illegal state latched）
        uErrInt     := 16#0005_0209;                // 0209 非法状态兜底（Illegal state fallback code）
        ePhase      := E_DL_TempBankPhase.eFault;   // 进终端安全态（Enter the terminal safe state）
END_CASE

(*------------------------------------------------------------------------------
 * 段 9｜复位（清故障、摘除状态与连续失败计数，温度保持供画面对比）
 *      Reset clears the fault, the drop state and the failure counters
 *-----------------------------------------------------------------------------*)
IF fbTrigReset.Q THEN
    bFaultLatch := FALSE;                       // 清故障锁存（Clear the fault latch）
    uErrInt     := 16#0000_0000;                // 清故障码（Clear the fault code）
    FOR i := 1 TO DL_DEV_MAX DO
        abDropped[i]     := FALSE;              // 清摘除标志（Clear the drop flag）
        anRecover[i]     := 0;                  // 清恢复计数（Clear the recovery counter）
        auCommFailCnt[i] := 0;                  // 清连续失败计数（Clear the failure counter）
    END_FOR
    uInfoCode := 16#0000_0000;                  // 复位当拍清信息码（Info code cleared on the reset cycle）
END_IF

(*------------------------------------------------------------------------------
 * 段 10｜出口映射与码位定级（单一优先级链，全拍只写一次 uErrorId）
 *      Outlet mapping with a single priority chain
 *-----------------------------------------------------------------------------*)
eState := ePhase;                               // 相位出口（Phase outlet）
bError := bFaultLatch;                          // 故障位只反映故障级锁存（Fault bit reflects the latch only）
IF bError THEN
    uErrorId := uErrInt;                        // 故障级码优先透出（Fault level code has priority）
ELSE
    uErrorId := uInfoCode;                      // 无故障透出本拍信息级码（Info code exposed otherwise）
END_IF
END_FUNCTION_BLOCK

(* ---- FB_DL_PumpPrimingSeq.st ---- *)
(*==============================================================================
 * 组件名称 (Component)  : FB_DL_PumpPrimingSeq
 * 所属子库 (Sublibrary) : DL_Process
 * 当前版本 (Version)    : 1.0.0
 * 兼容性   (Platform)   : CODESYS 3.5+ / TwinCAT 3 / 汇川 InoProShop / 施耐德 Machine Expert
 *                         仅依赖 Standard.library（TON / R_TRIG），零厂商私有库
 * 功能描述 (Function)   : 离心泵引水/自吸排气七态顺控：
 *                           eFill    开灌液阀：等 bFillValveFb 反馈，tFill 反馈超时 →
 *                                    eFault eCause=eFbFill；
 *                           eVent    开排气阀：等 bVentValveFb 反馈，tVent 反馈超时 →
 *                                    eFault eCause=eFbVent；
 *                           eConfirm 压力确认：fPrOutKpa >= fPrPrimeKpa → eDone（引水
 *                                    成功），tConfirm 窗内未达 → nRetries+1 回 eFill，
 *                                    nRetries > nRetryMax → eFault eCause=eNoPrime；
 *                           eRunning 主运态（本件只出态不接管泵启停）；eDone 引水确认
 *                                    完成，eRunning 下 bStop 正常停机 → eDone（引水序
 *                                    完成待复位），再 bStop/bReset → eIdle。
 *                         阀反馈超时各自 TON 段 0 刷新、分码 eFbFill/eFbVent（R190）。
 * 接口     (Interface)  : 输入 bStart/bStop/bReset、fPrOutKpa 泵出口压力（kPa）、
 *                         fPrPrimeKpa 引水成功判据（kPa）、bFillValveFb/bVentValveFb
 *                         阀反馈、tFill/tVent/tConfirm 各相窗、nRetryMax 重试上限；
 *                         输出 ePhase 七态、nRetries 重试计数、相指示 BOOL 组、bDone、
 *                         eCause、bError。
 * 边界     (Boundary)   : ① **属主边界（写死）：本件只管引水时序，不接管泵本体启停与
 *                         保护**（保护归 `FB_DL_PumpDryRunGuard` 族、主备切换归
 *                         `FB_DL_PumpChangeoverSeq`，三分域各管一段）。
 *                         ② 七态 CASE + ELSE 兜底 eFault（R6）；阀反馈/确认 TON 段 0
 *                         无条件刷新，IN 由当前相与反馈电平派生，无外部沿清零。
 *                         ③ 成因分码唯一（R190）：eFbFill / eFbVent / eNoPrime /
 *                         eNoData（压力非有限）/ eCfgIllegal。
 *                         ④ 组态闸：fPrPrimeKpa<=0、任一相时间 <= T#0S → 锁存 eFault
 *                         eCfgIllegal；**nRetryMax=0 为合法组态**（一次不过即故障）。
 *                         ⑤ 压力非有限 → eFault eNoData（R245）。
 *                         ⑥ bStop 在 eFault/eFill/eVent/eConfirm 中止回 eIdle；bStop 在
 *                         eRunning/eDone → eDone（正常停机完成态）；bReset 上升沿全清
 *                         nRetries（R311）。
 *                         ⑦ 零全局耦合（无 GVL / VAR_EXTERNAL / 物理地址）。
 * 分工声明 (Scope)      : 与 `FB_DL_PumpChangeoverSeq` 分工：引水启动 ≠ 主备切换；与
 *                         `FB_DL_PumpDryRunGuard`/`FB_DL_PumpDryRunProtect` 分工：引水
 *                         时序 ≠ 干转保护。
 * 来源标签 (Source Tag) : T2-2 ◐（LBP 工艺分层只借引水启动序分类事实，时序实现自研）
 * 码表     (Codes)      : 本件不占用任何全局数字码位。出口为 ENUM 七态 + UDINT 计数 +
 *                         BOOL 组 + ENUM 成因；数字码位待主控收口阶段统一派号。
 * 红线自检 (Redline)    : R1 ✓ 零 GVL/VAR_EXTERNAL ｜ R2 ✓ 零 %I/%Q/%M ｜ R3 ✓ 纯 IEC 61131-3
 *                         R4 ✓ 压力判据 >= 比较 + 非有限分码 + 组态闸 ｜ R5 ✓ 声明逐行同行双语注释
 *                         R6 ✓ 七态 CASE 含 ELSE ｜ R7 ✓ 三 TON/两 R_TRIG 段 0 无条件刷新
 * 修订历史 (Revision)   : 2026-11-20  v1.0.0  R48 首版（批次 4 · 序号 20）
 *                         验收向量：灌液阀反馈超时 → eFbFill；确认失败重试递增回 eFill；
 *                         nRetries > nRetryMax → eNoPrime；压力达标 → eDone → eRunning。
 *==============================================================================*)

TYPE E_DL_PpsPhase :
(
    eIdle    := 0,    // 待机 / Idle
    eFill    := 10,   // 灌液相 / Filling phase
    eVent    := 20,   // 排气相 / Venting phase
    eConfirm := 30,   // 压力确认相 / Pressure confirmation phase
    eRunning := 40,   // 主运态（只出态不接管泵启停）/ Main-run state
    eDone    := 50,   // 引水序完成（正常停机驻留）/ Priming sequence done
    eFault   := 90    // 故障（等复位）/ Fault, awaiting reset
);
END_TYPE

TYPE E_DL_PpsCause :
(
    eNone       := 0,   // 无异常 / No anomaly
    eCfgIllegal := 1,   // 组态非法 / Illegal configuration
    eNoData     := 2,   // 压力非有限 / Non-finite pressure
    eFbFill     := 3,   // 灌液阀反馈超时（R190 独立成因）/ Fill valve feedback timeout
    eFbVent     := 4,   // 排气阀反馈超时（R190 独立成因）/ Vent valve feedback timeout
    eNoPrime    := 5    // 重试耗尽未引水成功 / Retry budget exhausted, no prime
);
END_TYPE

FUNCTION_BLOCK FB_DL_PumpPrimingSeq
VAR_INPUT
    bStart       : BOOL := FALSE;   // 启动沿（eIdle 入灌液相） [-] / Start edge
    bStop        : BOOL := FALSE;   // 中止/停机（运行相回 eDone，其余回 eIdle） [-] / Stop
    bReset       : BOOL := FALSE;   // 复位，上升沿清全部锁存含 nRetries（R311） [-] / Reset, clears all latches
    fPrOutKpa    : LREAL := 0.0;    // 泵出口压力实测 [kPa] / Pump outlet pressure [kPa]
    fPrPrimeKpa  : LREAL := 150.0;  // 引水成功判据压力，域 > 0 [kPa] / Prime success pressure [kPa]
    bFillValveFb : BOOL := FALSE;   // 灌液阀开启反馈 [-] / Fill valve feedback
    bVentValveFb : BOOL := FALSE;   // 排气阀开启反馈 [-] / Vent valve feedback
    tFill        : TIME := T#10S;   // 灌液阀反馈超时窗，域 > T#0S [ms] / Fill feedback timeout [ms]
    tVent        : TIME := T#10S;   // 排气阀反馈超时窗，域 > T#0S [ms] / Vent feedback timeout [ms]
    tConfirm     : TIME := T#30S;   // 压力确认窗，域 > T#0S [ms] / Pressure confirm window [ms]
    nRetryMax    : UDINT := 3;      // 重试上限（=0 合法：一次不过即故障） [次] / Retry ceiling, 0 legal
END_VAR
VAR_OUTPUT
    ePhase      : E_DL_PpsPhase;    // 当前相出口 [-] / Present phase outlet
    nRetries    : UDINT;            // 引水重试计数出口 [次] / Retry count outlet
    bFillActive : BOOL;             // 灌液相指示（兼灌液阀命令参考） [-] / Fill phase indicator
    bVentActive : BOOL;             // 排气相指示（兼排气阀命令参考） [-] / Vent phase indicator
    bConfirmActive: BOOL;           // 压力确认相指示 [-] / Confirm phase indicator
    bRunning    : BOOL;             // 主运态指示 [-] / Main-run indicator
    bDone       : BOOL;             // 引水序完成指示 [-] / Priming done indicator
    eCause      : E_DL_PpsCause;    // 成因出口（锁存回放，R189） / Cause outlet, latched
    bError      : BOOL;             // 故障标志 [-] / Error flag
END_VAR
VAR
    _eState : E_DL_PpsPhase := E_DL_PpsPhase.eIdle;   // 内部相（CASE 唯一写入目标） / Internal phase
    _eCause : E_DL_PpsCause := E_DL_PpsCause.eNone;   // 成因锁存量 / Latched cause
    _bFault : BOOL;              // 故障锁存位（解除沿 = bReset 上升沿） / Latched fault bit
    _nRetry : UDINT := 0;        // 重试计数锁存量（bReset/bStop 全清） / Retry count latch
    _bNonFin: BOOL;              // 压力非有限当拍量 [-] / Non-finite pressure this scan
    _bCfgBad: BOOL;              // 组态非法当拍量 [-] / Illegal configuration this scan
    tonFbFill  : TON;            // 灌液阀反馈超时定时器，段 0 无条件调用 / Fill feedback timeout timer
    tonFbVent  : TON;            // 排气阀反馈超时定时器，段 0 无条件调用 / Vent feedback timeout timer
    tonConfirm : TON;            // 压力确认窗定时器，段 0 无条件调用 / Pressure confirm timer
    rtStart    : R_TRIG;         // 启动沿实例，段 0 无条件调用 / Start edge instance
    rtReset    : R_TRIG;         // 复位沿实例，段 0 无条件调用 / Reset edge instance
END_VAR
VAR CONSTANT
    DL_PPS_ZERO  : LREAL := 0.0;     // 非有限差值判零基准 [-] / Non-finite difference zero base
    DL_PPS_UDMAX : UDINT := 4294967295;   // UDINT 上限（重试计数饱和点） [次] / UDINT ceiling
END_VAR

(* —— 段 0：非有限判 + 组态闸 + 三 TON 两沿无条件周期刷新 —— *)
_bNonFin := (fPrOutKpa <> fPrOutKpa) OR ((fPrOutKpa - fPrOutKpa) <> DL_PPS_ZERO);   // 压力非有限（R245） / Non-finite pressure
_bCfgBad := (fPrPrimeKpa <= 0.0) OR (tFill <= T#0S) OR (tVent <= T#0S)
         OR (tConfirm <= T#0S);                         // 组态域闸（nRetryMax=0 合法不过闸） / Configuration gate
rtStart(CLK := bStart);                                 // 启动沿，每拍必调 / Start edge, every scan
rtReset(CLK := bReset);                                 // 复位沿，每拍必调 / Reset edge, every scan
tonFbFill(IN := (_eState = E_DL_PpsPhase.eFill) AND (NOT bFillValveFb), PT := tFill);    // 灌液反馈超时（反馈到即自复位） / Fill feedback timeout
tonFbVent(IN := (_eState = E_DL_PpsPhase.eVent) AND (NOT bVentValveFb), PT := tVent);    // 排气反馈超时 / Vent feedback timeout
tonConfirm(IN := (_eState = E_DL_PpsPhase.eConfirm), PT := tConfirm);   // 压力确认窗 / Pressure confirm window

(* —— 段 1：单拍量预清零（_eState/_eCause/_bFault/_nRetry 锁存量不入清单，R107） —— *)
bFillActive := FALSE;                                   // 灌液相指示预清 / Fill indicator preset
bVentActive := FALSE;                                   // 排气相指示预清 / Vent indicator preset
bConfirmActive := FALSE;                                // 确认相指示预清 / Confirm indicator preset
bRunning := FALSE;                                      // 主运指示预清 / Running preset
bDone := FALSE;                                         // 完成指示预清 / Done preset
bError := FALSE;                                        // 故障标志预清（R45 配对） / Error preset

(* —— 段 2：组态闸入故障 —— *)
IF _bCfgBad AND (NOT _bFault) THEN
    _bFault := TRUE;                                    // 锁存 / Latch
    _eCause := E_DL_PpsCause.eCfgIllegal;               // 归因：组态非法 / Cause: illegal config
    _eState := E_DL_PpsPhase.eFault;                    // 入故障相 / Enter fault
END_IF

(* —— 段 3：迁出链（bStop 分域语义 + bReset 全清 R311） —— *)
IF bStop AND (_eState <> E_DL_PpsPhase.eIdle) THEN
    IF (_eState = E_DL_PpsPhase.eRunning) OR (_eState = E_DL_PpsPhase.eDone) THEN
        _eState := E_DL_PpsPhase.eDone;                 // 运行/完成相停机 → eDone（正常停机完成态，头注释⑥） / Stop in run: to done
    ELSE
        IF _eState = E_DL_PpsPhase.eFault THEN
            _bFault := FALSE;                           // 停机优先清故障 / Stop wins over fault
            _eCause := E_DL_PpsCause.eNone;             // 清成因 / Clear cause
        END_IF
        _nRetry := 0;                                   // 中止全清重试计数（R311 同族） / Clear retries on abort
        _eState := E_DL_PpsPhase.eIdle;                 // 其余相中止回 eIdle / Abort to idle
    END_IF
END_IF
IF rtReset.Q THEN
    _bFault := FALSE;                                   // 清故障锁存（R311） / Clear fault latch
    _eCause := E_DL_PpsCause.eNone;                     // 清成因 / Clear cause
    _nRetry := 0;                                       // 复位沿全清重试计数（规格⑥） / Clear retries on reset edge
    _eState := E_DL_PpsPhase.eIdle;                     // 回待机 / Back to idle
END_IF

(* —— 段 4：七态顺控（只在无故障时推进；压力非有限 → eFault eNoData） —— *)
IF (NOT _bFault) AND (NOT _bCfgBad) AND (NOT bStop) THEN
    IF _bNonFin AND (_eState <> E_DL_PpsPhase.eIdle) AND (_eState <> E_DL_PpsPhase.eDone) THEN
        _bFault := TRUE;                                // 运行相压力非有限：故障锁存（规格⑤） / Non-finite in running phase
        _eCause := E_DL_PpsCause.eNoData;               // 归因分码：无有效数据 / Cause: no data
        _eState := E_DL_PpsPhase.eFault;                // 入故障相 / Enter fault
    ELSE
        CASE _eState OF

        E_DL_PpsPhase.eIdle:
            IF rtStart.Q THEN
                _nRetry := 0;                           // 新启动清重试计数 / Clear retries on new start
                _eState := E_DL_PpsPhase.eFill;         // 入灌液相 / Enter fill
            END_IF

        E_DL_PpsPhase.eFill:
            IF bFillValveFb THEN
                _eState := E_DL_PpsPhase.eVent;         // 灌液阀反馈到：进排气相 / Fill feedback: enter vent
            ELSIF tonFbFill.Q THEN
                _eCause := E_DL_PpsCause.eFbFill;       // 灌液反馈超时（R190 独立成因） / Fill feedback timeout
                _bFault := TRUE;                        // 锁存 / Latch
                _eState := E_DL_PpsPhase.eFault;        // 入故障相 / Enter fault
            END_IF

        E_DL_PpsPhase.eVent:
            IF bVentValveFb THEN
                _eState := E_DL_PpsPhase.eConfirm;      // 排气阀反馈到：进压力确认相 / Vent feedback: enter confirm
            ELSIF tonFbVent.Q THEN
                _eCause := E_DL_PpsCause.eFbVent;       // 排气反馈超时（R190 独立成因） / Vent feedback timeout
                _bFault := TRUE;                        // 锁存 / Latch
                _eState := E_DL_PpsPhase.eFault;        // 入故障相 / Enter fault
            END_IF

        E_DL_PpsPhase.eConfirm:
            IF fPrOutKpa >= fPrPrimeKpa THEN
                _eState := E_DL_PpsPhase.eRunning;      // 压力达标：转主运态（>= 判据禁浮点 =） / Pressure reached: to running
            ELSIF tonConfirm.Q THEN
                IF _nRetry < DL_PPS_UDMAX THEN
                    _nRetry := _nRetry + 1;             // 确认失败重试递增（饱和不回绕） / Increment retry, saturating
                END_IF
                IF _nRetry > nRetryMax THEN
                    _eCause := E_DL_PpsCause.eNoPrime;  // 重试耗尽（nRetryMax=0 时首轮即故障，合法） / Retry budget exhausted
                    _bFault := TRUE;                    // 锁存 / Latch
                    _eState := E_DL_PpsPhase.eFault;    // 入故障相 / Enter fault
                ELSE
                    _eState := E_DL_PpsPhase.eFill;     // 未耗尽：回灌液相重试 / Retry from fill
                END_IF
            END_IF

        E_DL_PpsPhase.eRunning:
            ;                                           // 主运驻留：本件只出态不接管泵启停（头注释①） / Held, pump control out of scope

        E_DL_PpsPhase.eDone:
            ;                                           // 完成驻留：由 bStop/bReset 迁出 / Held, exits via stop or reset

        E_DL_PpsPhase.eFault:
            ;                                           // 故障驻留：由迁出链处理 / Held by exit chain

        ELSE
            _eCause := E_DL_PpsCause.eCfgIllegal;       // 非法相位兜底归因 / Illegal phase cause
            _bFault := TRUE;                            // 锁存 / Latch
            _eState := E_DL_PpsPhase.eFault;            // 强拉故障相 / Force fault

        END_CASE
    END_IF
END_IF

(* —— 段 8：出口单点映射（相指示与相别同源，R191） —— *)
bFillActive := (_eState = E_DL_PpsPhase.eFill);         // 灌液相指示 / Fill indicator
bVentActive := (_eState = E_DL_PpsPhase.eVent);         // 排气相指示 / Vent indicator
bConfirmActive := (_eState = E_DL_PpsPhase.eConfirm);   // 确认相指示 / Confirm indicator
bRunning := (_eState = E_DL_PpsPhase.eRunning);         // 主运指示 / Running indicator
bDone := (_eState = E_DL_PpsPhase.eDone);               // 完成指示 / Done indicator
ePhase := _eState;                                      // 当前相出口 / Present phase outlet
nRetries := _nRetry;                                    // 重试计数出口 / Retry count outlet
eCause := _eCause;                                      // 成因出口 / Cause outlet
bError := _bFault OR _bCfgBad;                          // 故障标志 = 锁存或组态非法 / Error flag

END_FUNCTION_BLOCK

(* ---- FB_DL_R2rRunLogAudit.st ---- *)
(*==============================================================================
 * 组件名称 (Component)  : FB_DL_R2rRunLogAudit
 * 所属子库 (Sublibrary) : DL_Process
 * 当前版本 (Version)    : 1.0.0
 * 兼容性   (Platform)   : CODESYS 3.5+ / TwinCAT 3 / 汇川 InoProShop / 施耐德 Machine Expert
 *                         仅依赖 Standard.library（R_TRIG / LEN），零厂商私有库
 * 功能描述 (Function)   : R2R 调参批次审计算账。
 *                         把"谁在第几版改了哪些调参量"落成可追溯台账：每次提交沿到来时，
 *                         与上一份快照逐项比对，**只有真发生变化**才产生一条留痕记录（版本号 +1），
 *                         并把当时的参数值整组快照存档；未变化则不记账（防止操作员连点造成假账）。
 *                         三条固化纪律：
 *                           ① **变更沿留痕**：R_TRIG 段 0 无条件刷新；比对用"差值容差判等"
 *                              （浮点禁 =/<>，逐项 ABS 差 < fEps 视为同值）；
 *                           ② **台账计数饱和**：记录条数与版本号均以 UDINT 承载并在上限前
 *                              停止自增（饱和不回绕），饱和后置 bCntSaturated，绝不让计数回绕成小值；
 *                           ③ **快照缓冲满锁存**：缓冲深度满后拒记并锁存 bBufFull，
 *                              等运维导出台账后 bReset 清空重记，绝不静默丢账。
 *                         验收向量：
 *                           ① 首拍提交（基准快照）：版本 1，记录 1 条
 *                           ② 未改变任何参数再提交：版本不变、记录数不变、eNoChange（信息级）
 *                           ③ 只改第 3 项 +0.5：版本 2，记录 2 条，sLastTag = 本次标识
 *                           ④ 记录达深度 16 后再提交有变更：拒记 + bBufFull 锁存
 * 接口     (Interface)  : 入 bCommit 提交沿、sParamTag 参数组标识、afParam 当前调参量（1..8）、
 *                         nParamCnt 有效参数个数、fEps 判等容差、bReset 复位沿；
 *                         出 uLogCnt 台账条数、nRev 当前版本号、bChanged 记账脉冲（单拍）、
 *                         sLastTag 最近记账标识、bBufFull 缓冲满锁存、bCntSaturated 计数饱和标志、
 *                         eState 相、eCause 成因、bError 故障标志。
 * 边界     (Boundary)   : ① **属主边界（写死）：本件只做"调参快照 + 变更留痕 + 计数"，
 *                         不执行调参动作、不下发参数、不写 MES/磁盘**（分别属调参执行件与通讯件）；
 *                         ② **数组边界**：afParam 以字面量上界 8、缓冲以 16 声明（R104），
 *                         nParamCnt 与深度常量作运行时二次闸；
 *                         ③ **组态闸**：nParamCnt 须在 1..8、fEps 须 > 0，违反即锁存 eCfgIllegal；
 *                         ④ **计数饱和**：UDINT 上限前停止自增并置 bCntSaturated（饱和不回绕 R43 家族）；
 *                         ⑤ **非有限闸**：提交时任一参数非有限 → 拒记 + eParamBad（当拍，不锁存），
 *                         防止 NaN 污染台账信任根（R133）；
 *                         ⑥ **锁存解除式**：bBufFull 与 eFault 仅由 bReset 上升沿解除（R228B 唯一迁出）；
 *                         ⑦ 零全局耦合、零物理地址。
 * 分工声明 (Scope)      : 本件只管"调参审计台账"。不接管：调参算法执行
 *                         （属 FB_DL_R2rEwmaTuner）、参数合法性审查（属参数校验件）、
 *                         台账持久化（属 MES/文件件）。
 * 来源标签 (Source Tag) : ROADMAP 空勾真缺口 P1（R2R 调参审计，自研 clean-room）
 * 码表     (Codes)      : 本件不占用任何全局数字码位（零码位范式 R297）；诊断由 BOOL + ENUM 出口承担。
 * 红线自检 (Redline)    : R1 ✓ 零 GVL/VAR_EXTERNAL ｜ R2 ✓ 零 %I/%Q/%M ｜ R3 ✓ 纯 IEC 61131-3
 *                         R4 ✓ 数组闸 + 判等容差 + 计数饱和 + 非有限闸 ｜ R5 ✓ 声明逐行同行双语注释
 *                         R6 ✓ ENUM+CASE 含 ELSE 兜底 ｜ R7 ✓ R_TRIG 段 0 无条件刷新（本件无 TON）
 * 修订历史 (Revision)   : 2026-11-19  v1.0.0  R47 首版（批次 4 · 序号 17）
 *==============================================================================*)

TYPE ST_DL_RlaEntry :
STRUCT
    sTag   : STRING[15] := '';              // 参数组标识（≤15 字符） [-] / Parameter-group tag, up to 15 chars
    afVal  : ARRAY[1..8] OF LREAL;          // 记账时的参数值快照（1..8） [工程单位] / Parameter snapshot at logging time
    nCnt   : INT := 0;                      // 该条有效参数个数 [个] / Valid parameter count of this entry
    uRev   : UDINT := 0;                    // 该条对应版本号 [-] / Revision number of this entry
END_STRUCT
END_TYPE

TYPE E_DL_RlaState :
(
    eIdle  := 0,    // 待机相（等提交沿） / Idle, awaiting a commit edge
    eFault := 90    // 故障相（组态非法，等复位） / Fault, awaiting reset
);
END_TYPE

TYPE E_DL_RlaCause :
(
    eNone         := 0,   // 无异常 / No anomaly
    eFirstSnap    := 1,   // 首次基准快照（信息级） / First baseline snapshot, info level
    eNoChange     := 2,   // 提交但无变化（信息级，不记账） / Commit without change, info level
    eParamBad     := 3,   // 参数非有限（当拍拒记） / Non-finite parameter, rejected this scan
    eBufFull      := 4,   // 缓冲满（锁存，拒记） / Buffer full, latched, rejected
    eCfgIllegal   := 5,   // 组态非法（参数个数/容差越域） / Illegal configuration
    ePhaseBad     := 6    // 非法相位兜底 / Illegal phase fallback
);
END_TYPE

FUNCTION_BLOCK FB_DL_R2rRunLogAudit
VAR_INPUT
    bCommit   : BOOL := FALSE;         // 提交沿（记录一次调参结果） [-] / Commit edge, one audit record per edge
    sParamTag : STRING[15] := '';      // 参数组标识 [-] / Parameter-group tag
    afParam   : ARRAY[1..8] OF LREAL;  // 当前调参量（1..8） [工程单位] / Current parameter values, points 1..8
    nParamCnt : INT := 8;              // 有效参数个数，域 1..8 [个] / Valid parameter count, 1..8
    fEps      : LREAL := 1.0E-9;       // 判等容差，域 > 0 [工程单位] / Equality tolerance, > 0
    bReset    : BOOL := FALSE;         // 复位/清台账沿 [-] / Reset and clear edge
END_VAR
VAR_OUTPUT
    uLogCnt       : UDINT := 0;                          // 台账条数 [条] / Number of audit records
    nRev          : UDINT := 0;                          // 当前版本号 [-] / Current revision number
    bChanged      : BOOL := FALSE;                       // 记账脉冲（单拍） [-] / Logging pulse, single scan
    sLastTag      : STRING[15] := '';                    // 最近记账的参数组标识 [-] / Tag of the latest record
    bBufFull      : BOOL := FALSE;                       // 缓冲满锁存（等复位） [-] / Buffer full, latched
    bCntSaturated : BOOL := FALSE;                       // 计数饱和标志 [-] / Counter saturation flag
    eState        : E_DL_RlaState := E_DL_RlaState.eIdle;   // 相出口 [-] / Phase outlet
    eCause        : E_DL_RlaCause := E_DL_RlaCause.eNone;   // 成因出口（R190 归因唯一） [-] / Cause outlet
    bError        : BOOL := FALSE;                       // 故障标志（仅故障级成因） [-] / Error flag, fault level only
END_VAR
VAR
    _eState   : E_DL_RlaState := E_DL_RlaState.eIdle;    // 内部相（CASE 唯一写入目标） / Internal phase
    _eCause   : E_DL_RlaCause := E_DL_RlaCause.eNone;    // 成因锁存量 / Latched cause
    _bFault   : BOOL := FALSE;                           // 故障锁存位 / Latched fault bit
    _bBufFull : BOOL := FALSE;                           // 缓冲满锁存位 / Latched buffer-full bit
    _uCnt     : UDINT := 0;                              // 内部记录计数 / Internal record count
    _uRev     : UDINT := 0;                              // 内部版本号 / Internal revision number
    _bChanged : BOOL := FALSE;                           // 记账脉冲内部位（单拍） / Internal logging pulse
    _bInit    : BOOL := FALSE;                           // 基准快照已建立标志 / Baseline-established flag
    _bDiff    : BOOL := FALSE;                           // 本拍检出的差异标志 / Difference-found flag
    _bParamOk : BOOL := FALSE;                           // 参数有限性结论 / Parameter finiteness result
    _bCfgBad  : BOOL := FALSE;                           // 组态非法当拍量 / Illegal configuration this scan
    _i        : INT := 0;                                // 参数循环下标 / Parameter loop index
    _iIdx     : INT := 0;                                // 缓冲写指针（1..16） / Buffer write index
    afLast    : ARRAY[1..8] OF LREAL;                    // 上一版基准快照（1..8） / Previous baseline snapshot
    rtCommit  : R_TRIG;                                  // 提交沿实例，段 0 无条件调用 / Commit edge instance
    rtReset   : R_TRIG;                                  // 复位沿实例，段 0 无条件调用 / Reset edge instance
    astLog    : ARRAY[1..16] OF ST_DL_RlaEntry;          // 台账缓冲（深度字面量上界，R104） / Audit buffer
END_VAR
VAR CONSTANT
    DL_RLA_DEPTH  : UDINT := 16;         // 台账缓冲深度（与数组字面量上界同源） [条] / Audit buffer depth
    DL_RLA_PCNT   : INT := 8;            // 参数个数上限（与接口字面量上界同源） [个] / Parameter upper bound
    DL_RLA_NUM_MAX: UDINT := 16#FFFF_FFFE;  // 计数/版本饱和闸（留 1 个余量防回绕） [-] / Saturation gate
END_VAR

(* —— 段 0：组态闸 + 两沿无条件周期刷新（R228A；本件无 TON） —— *)
_bCfgBad := (nParamCnt < 1) OR (nParamCnt > DL_RLA_PCNT)                         // 参数个数须在 1..8 / Count within 1..8
         OR (fEps <= 0.0) OR (fEps <> fEps);                                     // 容差须为正且有限 / Tolerance positive and finite
rtCommit(CLK := bCommit);                                                        // 提交沿 / Commit edge
rtReset(CLK := bReset);                                                          // 复位沿 / Reset edge

(* —— 段 1：单拍量预清零（锁存量 _eCause/_bFault/_bBufFull/_uCnt/_uRev/_bInit 不入清单，R107） —— *)
_bChanged := FALSE;                                                              // 记账脉冲预清 / Logging pulse preset
_bDiff    := FALSE;                                                              // 差异标志预清 / Difference preset
bError    := FALSE;                                                              // 故障标志预清（R45 配对） / Error preset

(* —— 段 2：组态闸（非法即锁存） —— *)
IF _bCfgBad THEN
    _eCause := E_DL_RlaCause.eCfgIllegal;                                        // 归因：组态非法 / Cause: illegal configuration
    _bFault := TRUE;                                                             // 锁存 / Latch
    _eState := E_DL_RlaState.eFault;                                             // 入故障相 / Enter fault phase
END_IF

(* —— 段 3：迁出链（bReset 清双锁存并清台账；台账清空是运维显式动作） —— *)
IF rtReset.Q THEN
    _bFault   := FALSE;                                                          // 清故障锁存 / Clear fault latch
    _bBufFull := FALSE;                                                          // 清缓冲满锁存 / Clear the buffer-full latch
    _eCause   := E_DL_RlaCause.eNone;                                            // 清成因 / Clear cause
    _iIdx     := 1;                                                              // 写指针回 1 / Write index back to 1
    _uCnt     := 0;                                                              // 记录数清零 / Record count cleared
    _uRev     := 0;                                                              // 版本号清零 / Revision cleared
    _bInit    := FALSE;                                                          // 基准作废 / Baseline invalidated
    _eState   := E_DL_RlaState.eIdle;                                            // 回待机相 / Back to idle
END_IF

(* —— 段 4：相迁移（两相 CASE；故障相由段 3 迁出） —— *)
CASE _eState OF

E_DL_RlaState.eIdle:
    ;                                                                            // 待机相：记账在段 5 执行 / Logging happens in stage 5

E_DL_RlaState.eFault:
    ;                                                                            // 故障相：仅等复位 / Wait for the reset edge only

ELSE
    _eCause := E_DL_RlaCause.ePhaseBad;                                          // 归因：非法相位 / Cause: illegal phase
    _bFault := TRUE;                                                             // 锁存 / Latch
    _eState := E_DL_RlaState.eFault;                                             // 强拉故障相 / Force fault phase

END_CASE

(* —— 段 5：提交记账（有限性闸 → 差异比对 → 容量/饱和闸 → 落账） —— *)
IF (rtCommit.Q) AND (_eState = E_DL_RlaState.eIdle) AND (NOT _bCfgBad) THEN
    (* 有限性闸：任一有效参数非有限即当拍拒记（NaN 不得污染台账信任根，R133） *)
    _bParamOk := TRUE;                                                           // 结论初值 / Conclusion initial value
    FOR _i := 1 TO DL_RLA_PCNT DO
        IF _i <= nParamCnt THEN
            IF (afParam[_i] <> afParam[_i]) OR ((afParam[_i] - afParam[_i]) <> (afParam[_i] - afParam[_i])) THEN
                _bParamOk := FALSE;                                              // 检出非有限参数 / Non-finite parameter found
            END_IF
        END_IF
    END_FOR

    IF NOT _bParamOk THEN
        _eCause := E_DL_RlaCause.eParamBad;                                       // 归因：参数非有限 / Cause: non-finite parameter
    ELSIF NOT _bInit THEN
        (* 首次提交：建立基准快照并记第 1 条 *)
        IF _uCnt >= DL_RLA_DEPTH THEN
            _bBufFull := TRUE;                                                    // 容量闸（理论上首条不会满，仍显式判） / Capacity gate
            _eCause := E_DL_RlaCause.eBufFull;                                    // 归因：缓冲满 / Cause: buffer full
        ELSE
            FOR _i := 1 TO DL_RLA_PCNT DO
                afLast[_i] := afParam[_i];                                        // 建立基准 / Build the baseline
                astLog[_iIdx].afVal[_i] := afParam[_i];                           // 写记录值 / Write the record values
            END_FOR
            astLog[_iIdx].sTag := sParamTag;                                       // 写记录标识 / Write the record tag
            astLog[_iIdx].nCnt := nParamCnt;                                       // 写记录参数个数 / Write the record count
            _uRev := 1;                                                            // 版本号 1 / Revision 1
            astLog[_iIdx].uRev := _uRev;                                           // 记版本号 / Store the revision
            _uCnt := 1;                                                            // 记录数 1 / One record
            _iIdx := 2;                                                            // 写指针推进 / Advance the write index
            _bInit := TRUE;                                                        // 基准建立 / Baseline established
            _bChanged := TRUE;                                                     // 记账脉冲 / Logging pulse
            _eCause := E_DL_RlaCause.eFirstSnap;                                   // 归因：首次基准快照（信息级） / Cause: first baseline
        END_IF
    ELSE
        (* 差异比对：逐项差值容差判等，全部同值即"无变化" *)
        FOR _i := 1 TO DL_RLA_PCNT DO
            IF _i <= nParamCnt THEN
                IF ABS(afParam[_i] - afLast[_i]) > fEps THEN
                    _bDiff := TRUE;                                                // 检出差异 / Difference found
                END_IF
            END_IF
        END_FOR

        IF NOT _bDiff THEN
            _eCause := E_DL_RlaCause.eNoChange;                                    // 归因：无变化（信息级，不记账） / Cause: no change
        ELSIF _uCnt >= DL_RLA_DEPTH THEN
            _bBufFull := TRUE;                                                     // 缓冲满：锁存拒记 / Buffer full: latch and reject
            _eCause := E_DL_RlaCause.eBufFull;                                     // 归因：缓冲满 / Cause: buffer full
        ELSE
            FOR _i := 1 TO DL_RLA_PCNT DO
                afLast[_i] := afParam[_i];                                         // 更新基准 / Refresh the baseline
                astLog[_iIdx].afVal[_i] := afParam[_i];                            // 写记录值 / Write the record values
            END_FOR
            astLog[_iIdx].sTag := sParamTag;                                       // 写记录标识 / Write the record tag
            astLog[_iIdx].nCnt := nParamCnt;                                       // 写记录参数个数 / Write the record count
            IF _uRev < DL_RLA_NUM_MAX THEN
                _uRev := _uRev + 1;                                                // 版本号递增（饱和不回绕） / Revision increment
            ELSE
                bCntSaturated := TRUE;                                             // 版本号饱和 / Revision saturated
            END_IF
            astLog[_iIdx].uRev := _uRev;                                           // 记版本号 / Store the revision
            IF _uCnt < DL_RLA_NUM_MAX THEN
                _uCnt := _uCnt + 1;                                                // 记录数递增（饱和不回绕） / Count increment
            ELSE
                bCntSaturated := TRUE;                                             // 计数饱和 / Count saturated
            END_IF
            _iIdx := _iIdx + 1;                                                    // 写指针推进 / Advance the write index
            _bChanged := TRUE;                                                     // 记账脉冲 / Logging pulse
        END_IF
    END_IF
END_IF

(* —— 段 6：出口单点映射（名实双出口，R191） —— *)
uLogCnt       := _uCnt;                                                          // 记录数出口 / Record count outlet
nRev          := _uRev;                                                          // 版本号出口 / Revision outlet
bChanged      := _bChanged;                                                      // 记账脉冲出口 / Logging pulse outlet
sLastTag      := sParamTag;                                                      // 最近标识出口（与当拍提交同源） / Latest tag outlet
bBufFull      := _bBufFull;                                                      // 缓冲满出口 / Buffer-full outlet
eState        := _eState;                                                        // 相出口 / Phase outlet
eCause        := _eCause;                                                        // 成因出口 / Cause outlet
bError        := _bFault;                                                        // 故障标志 / Error flag

END_FUNCTION_BLOCK
